          def clipScaledValue(outputScaledValue, outputRange):
              if (outputRange[0] < outputRange[1]):
                  return clipWhenLowerLimitIsLessThanHigher(outputScaledValue, outputRange)
              else:
                  return clipWhenLowerLimitIsGreaterThanHigherLimit(outputScaledValue, outputRange)
              end
          end

          def clipWhenLowerLimitIsGreaterThanHigherLimit(outputScaledValue, outputRange):
              if (outputScaledValue < outputRange[1]):
                  return outputRange[1]
              elif (outputScaledValue > outputRange[0]):
                  return outputRange[0]
              else:
                  return outputScaledValue
              end
          end

          def clipWhenLowerLimitIsLessThanHigher(outputScaledValue, outputRange):
              if (outputScaledValue < outputRange[0]):
                  return outputRange[0]
              elif (outputScaledValue > outputRange[1]):
                  return outputRange[1]
              else:
                  return outputScaledValue
              end
          end

          slope = computeSlope(rawRange, scaledRange)
          intercept = computeIntercept(slope, rawRange, scaledRange)
          scaledValue = slope * value + intercept
          return clipScaledValue(scaledValue, scaledRange)
      end

      def limit(value, range):
          return scale(value, range, range)
      end


  rq_init_comm_if_connected(9, "1")
  rq_init_comm_if_connected(2, "2")
  rq_init_comm_if_connected(3, "3")
  rq_init_comm_if_connected(4, "4")
  rq_print_connected_grippers()
  rq_gripper_communication_thread = run rq_gripper_communication()
  set_closed_norm(97.6470588235294, "1")
  set_open_norm(1.1764705882352942, "1")
  set_closed_mm(0.0, "1")
  set_open_mm(53.0, "1")
  set_closed_norm(100.0, "2")
  set_open_norm(0.0, "2")
  set_closed_mm(0.0, "2")
  set_open_mm(50.0, "2")
  set_closed_norm(100.0, "3")
  set_open_norm(0.0, "3")
  set_closed_mm(0.0, "3")
  set_open_mm(50.0, "3")
  set_closed_norm(100.0, "4")
  set_open_norm(0.0, "4")
  set_closed_mm(0.0, "4")
  set_open_mm(50.0, "4")
  rq_current_limit_enabled = False
  while(not rq_gripper_communication_thread_started):
      sleep(0.008)
  end
  # end: URCap Installation Node
  step_count_b1809ffc_a9dc_407a_9cc4_7bc2f4a6af46 = 0.0
  thread Step_Counter_Thread_37d5f412_1517_4c3d_9382_b16793093957():
    while (True):
      step_count_b1809ffc_a9dc_407a_9cc4_7bc2f4a6af46 = step_count_b1809ffc_a9dc_407a_9cc4_7bc2f4a6af46 + 1.0
      sync()
    end
  end
  run Step_Counter_Thread_37d5f412_1517_4c3d_9382_b16793093957()
  global AMR_Position=struct(position_identifier=0, x1=0, x2=0, y1=0, y2=0, theta1=0, theta2=0)
  global CAM_Pose=p[0,0,0,0,0,0]
  global CAM_Relation=""
  global CMD_Abort=  False
  global CMD_Clear=  False
  global CMD_Reset=  False
  global CMD_Start=  False
  global CMD_Suspend=  False
  global CMD_Unhold=  False
  global CMD_Unsuspend=  False
  global CNT_Rack_Output=0
  global FNC_Freedrive=  False
  global PRC_TubCounter=0
  global STP=0
  global easyPickCount_4=0
  global easyPickCount_6=0
  global easyPickCount_7=0
  global easyPickCount_8=0
  global easyPickCount_9=0
  global easyPickNoObj_4=0
  global easyPickNoObj_6=0
  global easyPickNoObj_7=0
  global easyPickNoObj_8=0
  global easyPickNoObj_9=0
  global easyPickParts_4=0
  global easyPickParts_6=0
  global easyPickParts_7=0
  global easyPickParts_8=0
  global easyPickParts_9=0
  global Dosing_time=0
  global TMR_Barcode=0
  global Container_mid_1_p=p[-.379239199143, -.127191311915, .299999999998, .000000000046, -.000000000021, -1.247199999994]
  global Container_mid_1_q=[-2.477408934449926, -1.2969853503591224, -1.875639182904262, -1.539621866126728, 1.5731943360401213, -2.8009955944022717]
  global trigger_otw_p=p[-.364831738276, -.163967193938, .343299997821, .000000000046, -.000000000020, -1.148401333327]
  global trigger_otw_q=[-2.378283213085033, -1.2994862387706814, -1.7634300687554951, -1.6493302004167063, 1.573123683454141, -2.8011223671816943]
  global Waypoint_54_p=p[.008800512419, -.547926542621, .402696567415, -.589884378425, -.007228654778, -.061268144704]
  global Waypoint_54_q=[-1.2044575850116175, -1.3416667741588135, -1.8272563219070435, -0.9884541195682068, 1.3621035814285278, -2.7712565104113978]
  global Waypoint_77_p=p[-.178371829612, -.433927395311, .368082383916, -.086593488055, .704679941724, -.007869906074]
  global Waypoint_77_q=[-1.265390698109762, -1.3355963987163086, -1.7944865226745605, -1.7402602634825648, 0.8780410885810852, -2.7713127771960657]
  global Waypoint_83_p=p[.008800512419, -.547926542621, .402696567415, -.589884378425, -.007228654778, -.061268144704]
  global Waypoint_83_q=[-1.2044575850116175, -1.3416667741588135, -1.8272563219070435, -0.9884541195682068, 1.3621035814285278, -2.7712565104113978]
  global Waypoint_84_p=p[-.178371829612, -.433927395311, .368082383916, -.086593488055, .704679941724, -.007869906074]
  global Waypoint_84_q=[-1.265390698109762, -1.3355963987163086, -1.7944865226745605, -1.7402602634825648, 0.8780410885810852, -2.7713127771960657]
  global Vial_above_1_p=p[.017105793010, -.652093028359, .184920586844, .000000000272, .000000000270, 1.564063451276]
  global Vial_above_1_q=[-1.3375440709712851, -1.9618096977868804, -1.4665759083780685, -1.2837941559171444, 1.5732503672317195, -4.47276330421513]
  global Vial_pick_poi_1_p=p[.017105792852, -.648922724010, .093307568731, .000000000271, .000000000270, 1.564063451276]
  global Vial_pick_poi_1_q=[-1.3366329456391917, -2.0375277831965413, -1.6071432798879028, -1.0675084332049813, 1.57309887265915, -4.471135348858068]
  global Waypoint_86_p=p[.019227646885, -.648669633640, .184920586950, .000000000000, .000000000000, .024063451426]
  global Waypoint_86_q=[-1.3331129109407733, -1.9540750545686123, -1.4775914902901128, -1.280581784992414, 1.5733500744865856, -2.928303704452631]
  global Waypoint_87_p=p[-.032361834699, -.348336136197, .391475576335, -.000008499254, .000014589902, -.004651426820]
  global Waypoint_87_q=[-1.2709335019096129, -1.1914598663441005, -1.708995335060501, -1.8117888533498316, 1.5729683532263925, -2.8379347397710237]
  global Vial_3FG_plac_1_p=p[-.031858676359, -.349402499566, .145301120695, .000000000000, .000000000000, .000000000000]
  global Vial_3FG_plac_1_q=[-1.2723975525801707, -1.252376585823825, -2.3128114007049496, -1.1470592278900167, 1.5730548099411423, -2.8414815174610535]
  global Waypoint_88_p=p[-.032361834699, -.348336136197, .391475576335, -.000008499254, .000014589902, -.004651426820]
  global Waypoint_88_q=[-1.2709335019096129, -1.1914598663441005, -1.708995335060501, -1.8117888533498316, 1.5729683532263925, -2.8379347397710237]
  global cap_dump_1_p=p[-.139168676487, -.420163541420, .146096395183, .000000000000, .000000000000, .000000000000]
  global cap_dump_1_q=[-1.584588644510994, -1.5093464179777323, -2.1118449369620347, -1.091059703602438, 1.5728943834877336, -3.154014906686923]
  global Waypoint_89_p=p[-.032361834699, -.348336136197, .391475576335, -.000008499254, .000014589902, -.004651426820]
  global Waypoint_89_q=[-1.2709335019096129, -1.1914598663441005, -1.708995335060501, -1.8117888533498316, 1.5729683532263925, -2.8379347397710237]
  global Vial_3FG_plac_2_p=p[-.031858676359, -.349402499566, .145301120695, .000000000000, .000000000000, .000000000000]
  global Vial_3FG_plac_2_q=[-1.2723975525801707, -1.252376585823825, -2.3128114007049496, -1.1470592278900167, 1.5730548099411423, -2.8414815174610535]
  global Waypoint_90_p=p[-.032361834699, -.348336136197, .391475576335, -.000008499254, .000014589902, -.004651426820]
  global Waypoint_90_q=[-1.2709335019096129, -1.1914598663441005, -1.708995335060501, -1.8117888533498316, 1.5729683532263925, -2.8379347397710237]
  global cap_dump_2_p=p[-.139168676487, -.420163541420, .146096395183, .000000000000, .000000000000, .000000000000]
  global cap_dump_2_q=[-1.584588644510994, -1.5093464179777323, -2.1118449369620347, -1.091059703602438, 1.5728943834877336, -3.154014906686923]
  global Waypoint_91_p=p[-.032361834699, -.348336136197, .391475576335, -.000008499254, .000014589902, -.004651426820]
  global Waypoint_91_q=[-1.2709335019096129, -1.1914598663441005, -1.708995335060501, -1.8117888533498316, 1.5729683532263925, -2.8379347397710237]
  global Vial_liq_abov_1_p=p[-.025303660977, -.338758622354, .426628485936, -1.315858642253, .800043520260, -.928295855026]
  global Vial_liq_abov_1_q=[-0.3789628187762659, -1.5149522957256814, -2.263045310974121, 0.7870649534412841, -0.750984017048971, -3.2237566153155726]
  global Vial_liq_pick_3_p=p[-.002660428945, -.335984893034, .159389832934, -1.150456778400, .673175527684, -1.010612657503]
  global Vial_liq_pick_3_q=[-0.3660772482501429, -1.4503649038127442, -2.4056053161621094, -1.994692941705221, 0.8039668202400208, -0.2508929411517542]
  global Vial_liq_pick_4_p=p[-.041402486291, -.356791603314, .125395323246, -1.143483969075, .651070210027, -.878721885453]
  global Vial_liq_pick_4_q=[-0.4426233705502476, -1.437252121513727, -2.551930962114307, -1.776528229806984, 0.6562026234073748, -0.43018811960029524]
  global Vial_liq_abov_2_p=p[-.025303660977, -.338758622354, .426628485936, -1.315858642253, .800043520260, -.928295855026]
  global Vial_liq_abov_2_q=[-0.3789628187762659, -1.5149522957256814, -2.263045310974121, 0.7870649534412841, -0.750984017048971, -3.2237566153155726]
  global Liquid_midway_1_p=p[.057575295009, -.583081747994, .306414980749, -1.351675548728, .120935756539, -.096908606303]
  global Liquid_midway_1_q=[-0.895174805318014, -1.7035466633238734, -2.380953073501587, 0.631549521083496, 0.7706599235534668, -2.9455552736865442]
  global shake_3_p=p[.057574880217, -.583085370269, .306422893466, -1.360996190983, -.155555042453, -.438136255921]
  global shake_3_q=[-0.8951800505267542, -1.7035466633238734, -2.380937099456787, 0.6315542894550782, 0.7706599235534669, -2.5394540616517496]
  global shake_4_p=p[.057581636113, -.583090570002, .306439684073, -1.308767904323, .368530312677, .214926493520]
  global shake_4_q=[-0.8951714674579065, -1.7035395107665003, -2.380906343460083, 0.6315504747578125, 0.7706480026245118, -3.3161255787892268]
  global drop_above_3_p=p[.268235025993, -.467784390499, .226219872376, -1.027832627524, -.430841408251, 1.004603115937]
  global drop_above_3_q=[-0.935645882283346, -1.6663371525206507, -2.4252893924713135, 0.41966931402172847, 1.8470635414123535, -3.4600217978106897]
  global drop_above_4_p=p[.219042229014, -.470775657081, .133754190740, -.313004595901, -.344395319364, 1.500564994056]
  global drop_above_4_q=[-1.0601594887284795, -1.70046459045642, -2.0799996233759863, -0.7243227230676759, 1.9429634314685202, -4.115129153870795]
  global liq_tran_3_p=p[.213067510942, -.469567035397, .100231043184, .251862243732, .217902579404, 1.592812335393]
  global liq_tran_3_q=[-0.7789645168037476, -1.822364827406652, -1.8643518410805573, -1.252158963840138, 1.3768134449520435, -3.9328333233290254]
  global drop_above_5_p=p[.219042229014, -.470775657081, .133754190740, -.313004595901, -.344395319364, 1.500564994056]
  global drop_above_5_q=[-1.0601594887284795, -1.70046459045642, -2.0799996233759863, -0.7243227230676759, 1.9429634314685202, -4.115129153870795]
  global Waypoint_92_p=p[.187119460405, -.493959476151, .133754190608, -.313004596540, -.344395317757, 1.500564993991]
  global Waypoint_92_q=[-1.1418328121400876, -1.7310553375189475, -2.033634768766424, -0.772026910513711, 1.958578934631971, -4.201588449364511]
  global liq_tran_4_p=p[.195957706507, -.493022614126, .100231042689, .160718757180, .109807038912, 1.525321508623]
  global liq_tran_4_q=[-0.881740380645474, -1.8244526267589851, -1.865100964490387, -1.1608866323693583, 1.4631433601076713, -3.973915130363038]
  global drop_above_6_p=p[.219042229014, -.470775657081, .133754190740, -.313004595901, -.344395319364, 1.500564994056]
  global drop_above_6_q=[-1.0601594887284795, -1.70046459045642, -2.0799996233759863, -0.7243227230676759, 1.9429634314685202, -4.115129153870795]
  global drop_above_7_p=p[.268235025993, -.467784390499, .226219872376, -1.027832627524, -.430841408251, 1.004603115937]
  global drop_above_7_q=[-0.935645882283346, -1.6663371525206507, -2.4252893924713135, 0.41966931402172847, 1.8470635414123535, -3.4600217978106897]
  global Liquid_midway_2_p=p[.057575295009, -.583081747994, .306414980749, -1.351675548728, .120935756539, -.096908606303]
  global Liquid_midway_2_q=[-0.895174805318014, -1.7035466633238734, -2.380953073501587, 0.631549521083496, 0.7706599235534668, -2.9455552736865442]
  global Vial_drop_abo_1_p=p[.000324902251, -.648569523142, .221894115667, -.873462921366, 1.165852672573, -1.482720593185]
  global Vial_drop_abo_1_q=[-1.0576906334721352, -2.393016994184633, -0.9236232851859159, -2.5729213042279273, 0.7903331288549689, -0.33286325848155585]
  global Vial_liq_drop_1_p=p[.001020867953, -.647659915585, .092915870838, -.834762611599, 1.081942994823, -1.540647900176]
  global Vial_liq_drop_1_q=[-1.0631954168193474, -2.4447642951220825, -1.128811017825127, -2.1983115491972294, 0.8130148661460634, -0.38984988696911316]
  global Vial_drop_abo_2_p=p[.000324902251, -.648569523142, .221894115667, -.873462921366, 1.165852672573, -1.482720593185]
  global Vial_drop_abo_2_q=[-1.0576906334721352, -2.393016994184633, -0.9236232851859159, -2.5729213042279273, 0.7903331288549689, -0.33286325848155585]
  global pick_cont_otw_p=p[-.479450777041, .284140798427, .125270103493, -.276792173670, 2.098433187454, -2.121256516887]
  global pick_cont_otw_q=[-2.891505066548503, -1.9549266300590151, -2.231827259067863, -1.6654960117542226, 0.020810842514162875, -0.4019392172601952]
  global Powder_wayp1_p=p[-.472820924474, .292439826233, .207418370237, -.137787250486, 2.177332259632, -2.152029714756]
  global Powder_wayp1_q=[-2.911134078210732, -1.90240864358569, -1.968768330510411, -2.500365101593811, 0.11427687110891149, 0.0958980389250167]
  global Waypoint_2_p=p[-.357612884176, -.251084817998, .212379799667, -.858181193174, 1.714832512191, -1.687547565568]
  global Waypoint_2_q=[-1.620834863369681, -1.8936194567376496, -1.9821394403832038, -2.4599791457905273, 0.6296693672615152, 0.07625365420707819]
  global Decapp_above_1_p=p[-.013480295948, -.359153355979, .266194408367, -.879653555922, 1.646336924805, -1.709111068605]
  global Decapp_above_1_q=[-0.9632157249872035, -2.0163405763031657, -1.5968194594157152, -2.6579215719847085, 1.251243398585566, 0.047906446502667066]
  global Decapp_place_2_p=p[-.013480295890, -.359153356055, .160907502384, -.879653554902, 1.646336919740, -1.709111066456]
  global Decapp_place_2_q=[-0.9633402410919709, -2.1541179572356635, -1.6937729380888573, -2.4232786481058053, 1.2517342187662468, 0.04818402956922263]
  global Decapp_above_2_p=p[-.013480295948, -.359153355979, .266194408367, -.879653555922, 1.646336924805, -1.709111068605]
  global Decapp_above_2_q=[-0.9632157249872035, -2.0163405763031657, -1.5968194594157152, -2.6579215719847085, 1.251243398585566, 0.047906446502667066]
  global Waypoint_78_p=p[-.051450028091, -.519555688329, .365718563414, -1.287302938145, 1.077637394477, -1.218524965834]
  global Waypoint_78_q=[-0.9214276262416012, -1.8899696965062578, -1.4939326452510562, -2.840015661555725, 0.5585157189668353, 0.033997638875617575]
  global Decap_above_p=p[-.031863883354, -.349974838955, .288042264213, .000000000000, .000000000000, .000000000000]
  global Decap_above_q=[-1.271900116540503, -1.1670201114602632, -1.989291655468758, -1.5559360538518163, 1.573255119759632, -2.842476569674073]
  global Decapp_p=p[-.031864263150, -.349974612700, .230259377740, .000000000000, .000000000000, .000000000000]
  global Decapp_q=[-1.2723555431601419, -1.1810456878410935, -2.1291754890757737, -1.4020263844320349, 1.5732701843074919, -2.842325632263757]
  global Cap_above_p=p[-.224192409203, -.629599568633, .257274081142, .000015605575, -.000015166009, -1.647823825902]
  global Cap_above_q=[-1.710642681834492, -1.9674285251810462, -1.2705185053146897, -1.4742193161331247, 1.573506065067499, -1.6347709465008595]
  global Cap_place_p=p[-.224189049846, -.629597879697, .041885651757, .000015605572, -.000015166011, -1.647823825903]
  global Cap_place_q=[-1.7111696563854295, -2.13979870939016, -1.5941008764912503, -0.978265561728648, 1.5732789016410962, -1.6336328794662904]
  global OP_PowderA2_p=p[.009371277507, -.409434369247, .294169017766, -.823281033205, 1.709410851243, -1.698303593897]
  global OP_PowderA2_q=[-0.9994544761745754, -2.1395254572673217, -1.3437567783153916, -2.8143375616690456, 1.2617899549595724, 0.019614613715634555]
  global OP_PowderA_ab_1_p=p[-.012145216791, -.363335041455, .315325728178, -.777135478411, 1.752984823781, -1.740925591659]
  global OP_PowderA_ab_1_q=[-1.01634425044037, -2.024785947780374, -1.4658894155189923, -2.8070189735738786, 1.3091674480404514, 0.020022086766872782]
  global OP_PowderA_pick_p=p[-.019989579300, -.367909055381, .180100616111, -.546164737600, 1.935964719000, -1.930057109666]
  global OP_PowderA_pick_q=[-1.1609156816971709, -2.238534265251247, -1.4969295335038062, -2.556223512058769, 1.4532886345781417, 0.020741051754957773]
  global OP_PowderA_ab_2_p=p[-.012145216791, -.363335041455, .315325728178, -.777135478411, 1.752984823781, -1.740925591659]
  global OP_PowderA_ab_2_q=[-1.01634425044037, -2.024785947780374, -1.4658894155189923, -2.8070189735738786, 1.3091674480404514, 0.020022086766872782]
  global Op_PowA_wP_p=p[-.173727579245, -.372934016396, .295116627479, -.972390492433, 1.540962074418, -1.548745344994]
  global Op_PowA_wP_q=[-1.1740587397768483, -1.865656321049359, -1.7426943793777419, -2.679427276872525, 0.8588908769087338, 0.017944699631825187]
  global Waypoint_1_p=p[-.451048883256, -.340589460864, .308223661552, .097058877504, .091048998701, -1.578386010942]
  global Waypoint_1_q=[-2.222400490437643, -1.7554131946959437, -1.398173213005066, -1.6564461193480433, 1.5042352676391602, -2.2106884161578577]
  global Spatula_otw_p=p[-.222059999126, -.318140885971, .425288233229, -.000441582509, -.000128175490, 3.034387645854]
  global Spatula_otw_q=[-1.827769217553847, -1.3054220991219179, -1.546249130536875, -1.8605379988907114, 1.573101813278913, -0.15105460523915326]
  global pick_spat_L_abv_p=p[.239059466375, -.067212518441, .280720723617, .000017217488, -.000484427718, 3.106837214660]
  global pick_spat_L_abv_q=[0.292765616142962, -0.8565557553273315, -2.140199892763044, -1.715349495646084, 1.573623142106424, 1.8984976776985687]
  global spat_L_pick_p=p[.242468789885, -.067301915011, .193171208067, .000017217488, -.000484427718, 3.106837214657]
  global spat_L_pick_q=[0.2867414378807389, -0.8600077002089179, -2.3629148016312627, -1.4891831672860159, 1.5737695566221115, 1.8933890858591198]
  global spat_L_lift_p=p[.245402002494, -.067432373551, .289049296496, .000017217490, -.000484427724, 3.106837214657]
  global spat_L_lift_q=[0.2834351187564135, -0.8798320076811592, -2.1119436738532986, -1.7203314352121302, 1.573588313403067, 1.8891054681654005]
  global spat_L_side_p=p[.247133573905, -.017633681797, .289062935631, .000017217490, -.000484427724, 3.106837214657]
  global spat_L_side_q=[0.49719173575848863, -0.8582398211168538, -2.1182130454788215, -1.735610316654931, 1.5735817737572706, 2.1028402698705397]
  global spat_L_up_p=p[.247135508752, -.017665230822, .397130746165, .000017217490, -.000484427724, 3.106837214657]
  global spat_L_up_q=[0.49854946074076967, -0.9346239623559676, -1.808280269374471, -1.969158816463132, 1.5731020084036995, 2.1031742024348157]
  global spat_M_up_p=p[.245495561680, -.112112573515, .420343789747, .000026293989, -.000477463067, 3.067686800858]
  global spat_M_up_q=[0.09017908059107435, -1.0134242235449396, -1.71728844067247, -1.9814399845077446, 1.573013686840385, 1.733759055129931]
  global spat_M_pick_p=p[.244673518506, -.111985070134, .192299022723, .000026293990, -.000477463072, 3.067686800901]
  global spat_M_pick_q=[0.08834054082534859, -0.9272467647495475, -2.3438023910348154, -1.4411029496965373, 1.5736983399628084, 1.7342144371718433]
  global spat_S_Up_1_p=p[.252087445596, -.159242094834, .423281604617, .000026293954, -.000477463070, 3.067686800855]
  global spat_S_Up_1_q=[-0.09804692328730358, -1.0862987822056382, -1.6788706463996483, -1.9470242450550348, 1.5730147401359813, 1.5455107082823842]
  global spat_S_Pick_1_p=p[.245377020686, -.158668022535, .192285730279, .000026293985, -.000477463062, 3.067686800840]
  global spat_S_Pick_1_q=[-0.10087203759495189, -1.011188488703386, -2.311978084495874, -1.3890267520590838, 1.5735990551056096, 1.5450562970948172]
  global spat_S_Up_2_p=p[.252087445596, -.159242094834, .423281604617, .000026293954, -.000477463070, 3.067686800855]
  global spat_S_Up_2_q=[-0.09804692328730358, -1.0862987822056382, -1.6788706463996483, -1.9470242450550348, 1.5730147401359813, 1.5455107082823842]
  global spat_flatM_up_p=p[.229022666361, -.211442909333, .418634047126, .000026293953, -.000477463083, 3.067686800888]
  global spat_flatM_up_q=[-0.30183372580416545, -1.1157042924275036, -1.6775646144685776, -1.9189678841796578, 1.5730340557943228, 1.341766142011193]
  global spat_flatM_pick_p=p[.241028983327, -.208057297586, .192270533170, .000026293950, -.000477463079, 3.067686800885]
  global spat_flatM_pick_q=[-0.2805687960562633, -1.1003763929487214, -2.271431297337675, -1.3404236887924883, 1.5734924238720627, 1.3653813047742556]
  global spat_flatS_up_p=p[.237651953780, -.253943828614, .403961222825, .000026293950, -.000477463092, 3.067686800841]
  global spat_flatS_up_q=[-0.42363550926974103, -1.1939944599502539, -1.6745915127240307, -1.843675057902054, 1.5731001874678698, 1.220082820532415]
  global spat_flatS_pick_p=p[.241325662334, -.251726327528, .192256842740, .000026293947, -.000477463087, 3.067686800841]
  global spat_flatS_pick_q=[-0.4144907797170738, -1.1967447109013012, -2.21926362252748, -1.2962499335425761, 1.5733885098427622, 1.2314402238866728]
  global spat_S_pick_p=p[.238158866340, -.157926795425, .192632100345, .000026293989, -.000477463069, 3.067686800857]
  global spat_S_pick_q=[-0.10084756991493293, -0.9881392730064915, -2.3204232610157494, -1.403630829593915, 1.5736254260650586, 1.5450653591083503]
  global spat_S_up_p=p[.244260523725, -.164466690315, .417087579736, .000026293988, -.000477463072, 3.067686800857]
  global spat_S_up_q=[-0.12101499604198729, -1.0718307017854336, -1.7023391702814736, -1.938028805938881, 1.573044424728474, 1.5226045951991447]
  global spat_S_Up_3_p=p[.252087445596, -.159242094834, .423281604617, .000026293954, -.000477463070, 3.067686800855]
  global spat_S_Up_3_q=[-0.09804692328730358, -1.0862987822056382, -1.6788706463996483, -1.9470242450550348, 1.5730147401359813, 1.5455107082823842]
  global spat_S_Pick_2_p=p[.245377020686, -.158668022535, .192285730279, .000026293985, -.000477463062, 3.067686800840]
  global spat_S_Pick_2_q=[-0.10087203759495189, -1.011188488703386, -2.311978084495874, -1.3890267520590838, 1.5735990551056096, 1.5450562970948172]
  global spat_S_Up_4_p=p[.252087445596, -.159242094834, .423281604617, .000026293954, -.000477463070, 3.067686800855]
  global spat_S_Up_4_q=[-0.09804692328730358, -1.0862987822056382, -1.6788706463996483, -1.9470242450550348, 1.5730147401359813, 1.5455107082823842]
  global PosA_up_p=p[.016801192651, -.634607931192, .234972649145, -1.090660933959, 1.404791542935, -1.413645191218]
  global PosA_up_q=[-1.0269853941957567, -2.5566815932087046, -0.7524196965257657, -2.981505396440104, 0.8113680441070815, 0.02148045637209592]
  global PosA_pick_p=p[.015038978729, -.636805282702, .098001171702, -1.090660933960, 1.404791542941, -1.413645191214]
  global PosA_pick_q=[-1.030538681681108, -2.6868026737636344, -0.8591268496433386, -2.7445819191995, 0.8086593798745287, 0.021358164952170952]
  global trigger_otw_2_p=p[-.364831738276, -.163967193938, .343299997821, .000000000046, -.000000000020, -1.148401333327]
  global trigger_otw_2_q=[-2.378283213085033, -1.2994862387706814, -1.7634300687554951, -1.6493302004167063, 1.573123683454141, -2.8011223671816943]
  global Postions_otw_p=p[-.010896578244, -.533368729951, .288851175116, -1.233738470894, 1.195331112012, -1.207314088469]
  global Postions_otw_q=[-0.898791023514228, -2.078490033037677, -1.4499891355755317, -2.7624416226992476, 0.6570218891920963, 0.02136606178275929]
  global spat_S_Up_5_p=p[.252087445596, -.159242094834, .423281604617, .000026293954, -.000477463070, 3.067686800855]
  global spat_S_Up_5_q=[-0.09804692328730358, -1.0862987822056382, -1.6788706463996483, -1.9470242450550348, 1.5730147401359813, 1.5455107082823842]
  global spat_S_Pick_3_p=p[.245377020686, -.158668022535, .192285730279, .000026293985, -.000477463062, 3.067686800840]
  global spat_S_Pick_3_q=[-0.10087203759495189, -1.011188488703386, -2.311978084495874, -1.3890267520590838, 1.5735990551056096, 1.5450562970948172]
  global spat_S_Up_6_p=p[.252087445596, -.159242094834, .423281604617, .000026293954, -.000477463070, 3.067686800855]
  global spat_S_Up_6_q=[-0.09804692328730358, -1.0862987822056382, -1.6788706463996483, -1.9470242450550348, 1.5730147401359813, 1.5455107082823842]
  global spat_S_Up_7_p=p[.252087445596, -.159242094834, .423281604617, .000026293954, -.000477463070, 3.067686800855]
  global spat_S_Up_7_q=[-0.09804692328730358, -1.0862987822056382, -1.6788706463996483, -1.9470242450550348, 1.5730147401359813, 1.5455107082823842]
  global spat_S_Pick_4_p=p[.245377020686, -.158668022535, .192285730279, .000026293985, -.000477463062, 3.067686800840]
  global spat_S_Pick_4_q=[-0.10087203759495189, -1.011188488703386, -2.311978084495874, -1.3890267520590838, 1.5735990551056096, 1.5450562970948172]
  global spat_S_Up_8_p=p[.252087445596, -.159242094834, .423281604617, .000026293954, -.000477463070, 3.067686800855]
  global spat_S_Up_8_q=[-0.09804692328730358, -1.0862987822056382, -1.6788706463996483, -1.9470242450550348, 1.5730147401359813, 1.5455107082823842]
  global PosB_up_p=p[.239472634782, -.492481416782, .220767759213, -1.233738470883, 1.195331111998, -1.207314088469]
  global PosB_up_q=[-0.5800230603397054, -2.4076296700885997, -1.0699783327330836, -2.8116344407747427, 0.9750472858169287, 0.017627507888886562]
  global PosB_pick_p=p[.240630296955, -.494558620171, .096392895280, -1.233740573549, 1.195309876041, -1.207293779132]
  global PosB_pick_q=[-0.5816146260408139, -2.553273721769836, -1.1376320925804277, -2.5983292591462153, 0.9740936784345416, 0.017625262979849232]
  global PosC_up_p=p[.241566602786, -.359249123455, .230260583862, -1.233738470888, 1.195331111997, -1.207314088449]
  global PosC_up_q=[-0.39573787962534546, -2.2019009616581497, -1.4115270142506517, -2.675987785326166, 1.160180741930842, 0.01687917643039505]
  global PosC_pick_p=p[.240633854030, -.361553124916, .093979792658, -1.233738470878, 1.195331111997, -1.207314088469]
  global PosC_pick_q=[-0.39992427526118757, -2.386042391328985, -1.4894374567278712, -2.414022930893381, 1.1566786195951169, 0.01712017454263659]
  global Pow_decap_up_p=p[-.017556487132, -.367519866742, .275835445416, -.605635182849, 1.892518157522, -1.890848751165]
  global Pow_decap_up_q=[-1.1272088681128203, -2.1173924123331025, -1.4250048354055203, -2.7485980486387676, 1.4193896902217862, 0.023247957637719453]
  global pow_decap_place_p=p[-.020433194420, -.368310202914, .161281291611, -.605635182838, 1.892518157522, -1.890848751163]
  global pow_decap_place_q=[-1.132360890531647, -2.2521863255983092, -1.5302136899970318, -2.5086176644751683, 1.4149282844269635, 0.02347140074572661]
  global Decap_up_p=p[-.018339217391, -.367674469480, .249553854268, -.546164737599, 1.935964719000, -1.930057109666]
  global Decap_up_q=[-1.158124747223252, -2.1569920012936787, -1.4340832185069745, -2.7006032680036753, 1.4556626828962336, 0.02060977878679182]
  global Decap_pick_p=p[-.020429098827, -.367971872627, .161604333799, -.546164737600, 1.935964719000, -1.930057109666]
  global Decap_pick_q=[-1.161653098289774, -2.263509236689538, -1.5087211318402236, -2.519459740767391, 1.452646640403743, 0.02077912034002202]
  global spat_S_Up_9_p=p[.252087445596, -.159242094834, .423281604617, .000026293954, -.000477463070, 3.067686800855]
  global spat_S_Up_9_q=[-0.09804692328730358, -1.0862987822056382, -1.6788706463996483, -1.9470242450550348, 1.5730147401359813, 1.5455107082823842]
  global spat_S_Pick_5_p=p[.245377020686, -.158668022535, .192285730279, .000026293985, -.000477463062, 3.067686800840]
  global spat_S_Pick_5_q=[-0.10087203759495189, -1.011188488703386, -2.311978084495874, -1.3890267520590838, 1.5735990551056096, 1.5450562970948172]
  global spat_S_Up_10_p=p[.252087445596, -.159242094834, .423281604617, .000026293954, -.000477463070, 3.067686800855]
  global spat_S_Up_10_q=[-0.09804692328730358, -1.0862987822056382, -1.6788706463996483, -1.9470242450550348, 1.5730147401359813, 1.5455107082823842]
  global Cap_Pos1_up_p=p[-.009204590651, -.630414532143, .209553215594, .000015605636, -.000015165972, -1.647823825918]
  global Cap_Pos1_up_q=[-1.3712235360848153, -1.8956436160717116, -1.4937179908129403, -1.3227667547680468, 1.5734078303557693, -1.294583528806303]
  global Cap_pos1_p=p[-.009202676635, -.630420568421, .169124041327, .000015605637, -.000015165972, -1.647823825918]
  global Cap_pos1_q=[-1.3713472255781163, -1.9233675297983162, -1.5632855513360973, -1.2254750650219144, 1.573366428933177, -1.2943660310427454]
  global Cap_Pos2_up_p=p[.211716053312, -.494057775376, .215280069366, .000015605634, -.000015165975, -1.647823825915]
  global Cap_Pos2_up_q=[-0.9145242936692304, -1.674696899505042, -1.7522162453415309, -1.2851708271213624, 1.5732187144557628, -0.8372657504386876]
  global Cap_Pos2_p=p[.212489912868, -.496566704351, .174147693321, .000015605636, -.000015165975, -1.647823825915]
  global Cap_Pos2_q=[-0.9164207524863208, -1.713567851985026, -1.8189683536262713, -1.1795477490971313, 1.5731464491112233, -0.8388186043721344]
  global Cap_Pos3_up_p=p[.215414026072, -.362498267015, .204704869421, .000015605620, -.000015165977, -1.647823825911]
  global Cap_Pos3_up_q=[-0.7126949721702758, -1.3944102858194336, -2.0491785338653417, -1.268480216466319, 1.5731602525658304, -0.6347529509142049]
  global Cap_pos3_p=p[.215414769079, -.362497999431, .173969495144, .000015605637, -.000015165975, -1.647823825916]
  global Cap_pos3_q=[-0.7128543668961971, -1.4224209260451453, -2.1096401714367516, -1.1800078429832341, 1.573077069822543, -0.6346164729408441]
  global Dosing_time_is_counting=False
  global TMR_Barcode_is_counting=False
  thread Timer_Thread():
    while (True):
      if (Dosing_time_is_counting):
        Dosing_time = Dosing_time + get_steptime()
      end
      if (TMR_Barcode_is_counting):
        TMR_Barcode = TMR_Barcode + get_steptime()
      end
      sync()
    end
  end
  run Timer_Thread()
  def Sub_Vision_V18():
    $ 817 "Sub_Vision_V18" "noBreak"
    $ 818 "PreSettings"
    $ 819 "CAM_LM_Detected≔ False "
    global CAM_LM_Detected=  False
    $ 820 "CAM_Captures≔0"
    global CAM_Captures=0
    $ 821 "CAM_Pose≔p[0,0,0,0,0,0]"
    global CAM_Pose=p[0,0,0,0,0,0]
    $ 822 "CAM_LM_Refinmnt≔ False "
    global CAM_LM_Refinmnt=  False
    $ 823 "CAM_LM_Refined≔ False "
    global CAM_LM_Refined=  False
    $ 824 "CAM_LM_Deviatn≔p[0,0,0,0,0,0]"
    global CAM_LM_Deviatn=p[0,0,0,0,0,0]
    $ 825 "CAM_LM_ID≔0"
    global CAM_LM_ID=0
    $ 826 "CAM_Done≔ False "
    global CAM_Done=  False
    $ 827 "CAM_CNT_Obj≔0"
    global CAM_CNT_Obj=0
    $ 828 "CAM_Result = []"
    CAM_Result = []
    $ 829 "OBJ_Detected≔ False "
    global OBJ_Detected=  False
    $ 830 "FRM_Reference≔p[0,0,0,0,0,0]"
    global FRM_Reference=p[0,0,0,0,0,0]
    $ 831 "'=========='"
    # '=========='
    $ 832 "Switch Action"
    switch_1 = Action
    $ 833 "Case 13"
    if (13 == switch_1):
    elif (15 == switch_1):
      $ 951 "Case 15"
    elif (131 == switch_1):
      $ 997 "Case 131"
      $ 998 "Read (SensoPart)"
      $ 999 "Action_Info≔'search for landmark'"
      global Action_Info="search for landmark"
      $ 1000 "CAM_LM≔CAM_LMs[4]"
      global CAM_LM=CAM_LMs[4]
      $ 1001 "CAM_Relation≔CAM_LM.capture_relation"
      global CAM_Relation=CAM_LM.capture_relation
      $ 1002 "go to capture pose"
      $ 1005 "If ITM_ID≟1 and JIG≟7"
      if (ITM_ID == 1  and  JIG == 7):
        $ 1006 "PSE_T≔uLM_Cap_SSRack"
        global PSE_T=uLM_Cap_SSRack
      else:
        $ 1007 "ElseIf ITM_ID≟5 and JIG≟7"
        if (ITM_ID == 5  and  JIG == 7):
          $ 1008 "PSE_T≔FRM_Cap_SSRack"
          global PSE_T=FRM_Cap_SSRack
        else:
          $ 1011 "ElseIf ITM_ID≟1 and JIG≟15"
          if (ITM_ID == 1 and JIG == 15):
            $ 1012 "MoveJ"
            $ 1013 "Container_mid_1" "breakAfter"
            movej(get_inverse_kin(Container_mid_1_p, qnear=Container_mid_1_q), a=1.3962634015954636, v=1.0471975511965976, r=0.05)
            $ 1015 "PSE_T≔FRM_Container_const"
            global PSE_T=p[-0.5003348223692186,0.35061804815168285,0.41579001388808423,-5.092943187272062E-5,1.0145185065363121E-4,-2.764319258713288]
          else:
            $ 1016 "ElseIf ITM_ID≟1 and JIG≟21"
            if (ITM_ID == 1 and JIG == 21):
              $ 1017 "PSE_T≔FRM_PoTS_const"
              global PSE_T=p[-0.5306792777448894,-0.11733736113273928,0.4723291514857741,-1.2750528643267135E-5,1.622694849249343E-6,-2.208498084105121]
            else:
              $ 1018 "ElseIf ITM_ID≟1 and JIG≟17"
              if (ITM_ID == 1 and JIG == 17):
                $ 1019 "MoveJ"
                $ 1020 "trigger_otw" "breakAfter"
                movej(get_inverse_kin(trigger_otw_p, qnear=trigger_otw_q), a=1.3962634015954636, v=1.0471975511965976, r=0.05)
                $ 1021 "PSE_T≔FRM_weigh_scale_const"
                global PSE_T=p[-0.3552030492367321,0.06852934966463993,0.4723405535118315,-1.0342323845904682E-4,-1.3726098069249118E-5,-2.169178331189411]
              end
            end
          end
        end
      end
      $ 1022 "do_transition(PSE_T, keep_rxry=False)"
      do_transition(PSE_T, keep_rxry=False)
      $ 1023 "Set"
      set_tcp(p[0.0,0.0,0.161,3.1415,0.0,0.0])
      $ 1024 "MoveJ"
      $ 1025 "PSE_T" "breakAfter"
      movej(PSE_T, a=1.3962634015954636, v=1.7453292519943295)
      $ 1026 "CAM_Pose≔get_actual_tcp_pose()"
      global CAM_Pose= get_actual_tcp_pose ()
      $ 1027 "Loop  not CAM_Done and  not ERROR.FLAG and  not CMD_Stop"
      while (  not  CAM_Done  and    not  ERROR.FLAG  and    not  CMD_Stop):
        $ 1028 "adjust capture pose"
        $ 1029 "If CAM_LM_Detected and CAM_LM_Refinmnt"
        if (CAM_LM_Detected  and  CAM_LM_Refinmnt):
          $ 1030 "PSE_T≔p[0,0,0.300,0,0,0]"
          global PSE_T=p[0,0,0.300,0,0,0]
          $ 1031 "CAM_Pose≔PSE_T"
          global CAM_Pose=PSE_T
          $ 1032 "If  not is_reachable(FRM_Reference,[PSE_T])"
          if (  not  is_reachable(FRM_Reference,[PSE_T])):
            $ 1033 "Error"
            $ 1034 "set_error(ERROR_POSE_NOT_REACHABLE)"
            set_error(ERROR_POSE_NOT_REACHABLE)
          end
          $ 1035 "If  not ERROR.FLAG"
          if (  not  ERROR.FLAG):
            $ 1036 "MoveJ"
            $ 1037 "PSE_T" "breakAfter"
            set_tcp(p[0.0,0.0,0.161,0.0,0.0,0.0])
            movej(pose_trans(FRM_Reference, PSE_T), a=0.8726646259971648, v=1.3962634015954636)
            $ 1038 "CAM_LM_Refined≔ True "
            global CAM_LM_Refined=  True
          end
        else:
          $ 1039 "ElseIf  not CAM_LM_Detected and CAM_Captures>0"
          if (  not  CAM_LM_Detected  and  CAM_Captures>0):
            $ 1040 "MoveL"
            $ 1041 "If FRM_Reference≟p[0,0,0,0,0,0]"
            if (FRM_Reference == p[0,0,0,0,0,0]):
              $ 1042 "PSE_T≔get_random_pose(pose_ref=CAM_Pose, mode='cubic', range_max=[0.150,0.150,0.015])"
              global PSE_T=get_random_pose(pose_ref=CAM_Pose, mode="cubic", range_max=[0.150,0.150,0.015])
            else:
              $ 1047 "Else" "noBreak"
              $ 1048 "PSE_T≔get_random_pose(pose_ref=CAM_Pose, mode='rotation', range_max=[10,10,0])"
              global PSE_T=get_random_pose(pose_ref=CAM_Pose, mode="rotation", range_max=[10,10,0])
              $ 1049 "CAM_LM_Refined≔ True "
              global CAM_LM_Refined=  True
            end
            $ 1050 "If get_inverse_kin_has_solution(pose_trans(FRM_Reference, PSE_T))"
            if (get_inverse_kin_has_solution( pose_trans (FRM_Reference, PSE_T))):
              $ 1051 "Comment"
              # Comment
              $ 1052 "PSE_T" "breakAfter"
              set_tcp(p[0.0,0.0,0.161,3.1415,0.0,0.0])
              movel(pose_trans(FRM_Reference, PSE_T), a=0.03, v=0.05)
            else:
              $ 1053 "Else" "noBreak"
              $ 1054 "'If random pose is out of reach, set the initial cam pose'"
              # 'If random pose is out of reach, set the initial cam pose'
              $ 1055 "PSE_T≔CAM_Pose"
              global PSE_T=CAM_Pose
            end
          end
        end
        $ 1056 "Wait: 2.0"
        sleep(2.0)
        $ 1057 "trigger"
        $ 1058 "If ITM_ID≟1 and JIG≟7"
        if (ITM_ID == 1  and  JIG == 7):
          # begin: URCap Program Node
          #   Source: SensoPart VISOR Robotic, 2.0.6, SensoPart Industriesensorik GmbH
          #   Type: VISOR Trigger
          $ 1059 "# 1 VISOR Trigger"
          visor_changeJob(1, "Landmark_INVITE_2", 6000)
          visor_trigger(1, 6000, "arm")
          # end: URCap Program Node
        else:
          $ 1060 "ElseIf ITM_ID≟5 and JIG≟7"
          if (ITM_ID == 5  and  JIG == 7):
            # begin: URCap Program Node
            #   Source: SensoPart VISOR Robotic, 2.0.6, SensoPart Industriesensorik GmbH
            #   Type: VISOR Trigger
            $ 1061 "# 1 VISOR Trigger"
            visor_changeJob(1, "Landmark_INVITE_2", 6000)
            visor_trigger(1, 6000, "arm")
            # end: URCap Program Node
          else:
            $ 1062 "ElseIf ITM_ID≟13 and JIG≟7"
            if (ITM_ID == 13  and  JIG == 7):
              # begin: URCap Program Node
              #   Source: SensoPart VISOR Robotic, 2.0.6, SensoPart Industriesensorik GmbH
              #   Type: VISOR Trigger
              $ 1063 "# 1 VISOR Trigger"
              visor_changeJob(1, "Landmark_INVITE_2", 6000)
              visor_trigger(1, 6000, "arm")
              # end: URCap Program Node
            else:
              $ 1064 "ElseIf ITM_ID≟1 and JIG≟15"
              if (ITM_ID == 1 and JIG == 15):
                # begin: URCap Program Node
                #   Source: SensoPart VISOR Robotic, 2.0.6, SensoPart Industriesensorik GmbH
                #   Type: VISOR Trigger
                $ 1065 "# 1 VISOR Trigger"
                visor_changeJob(1, "QR_box", 6000)
                visor_trigger(1, 6000, "arm")
                # end: URCap Program Node
              else:
                $ 1066 "ElseIf ITM_ID≟1 and JIG≟21"
                if (ITM_ID == 1 and JIG == 21):
                  # begin: URCap Program Node
                  #   Source: SensoPart VISOR Robotic, 2.0.6, SensoPart Industriesensorik GmbH
                  #   Type: VISOR Trigger
                  $ 1067 "# 1 VISOR Trigger"
                  visor_changeJob(1, "PoTS", 6000)
                  visor_trigger(1, 6000, "arm")
                  # end: URCap Program Node
                else:
                  $ 1068 "ElseIf ITM_ID≟1 and JIG≟17"
                  if (ITM_ID == 1 and JIG == 17):
                    # begin: URCap Program Node
                    #   Source: SensoPart VISOR Robotic, 2.0.6, SensoPart Industriesensorik GmbH
                    #   Type: VISOR Trigger
                    $ 1069 "# 1 VISOR Trigger"
                    visor_changeJob(1, "Weigh_target", 6000)
                    visor_trigger(1, 6000, "arm")
                    # end: URCap Program Node
                  end
                end
              end
            end
          end
        end
        $ 1073 "TM_3D_Found≔visor_partsFound(1)"
        global TM_3D_Found= visor_partsFound (1)
        $ 1074 "If TM_3D_Found>0"
        if (TM_3D_Found>0):
          $ 1075 "CAM_LM_Detected≔ True "
          global CAM_LM_Detected=  True
          $ 1076 "CAM_Captures≔0"
          global CAM_Captures=0
        else:
          $ 1077 "Else" "noBreak"
          $ 1078 "CAM_LM_Detected≔ False "
          global CAM_LM_Detected=  False
          $ 1079 "CAM_Captures≔CAM_Captures+1"
          global CAM_Captures=CAM_Captures+1
        end
        $ 1084 "result"
        $ 1085 "If CAM_LM_Detected"
        if (CAM_LM_Detected):
          $ 1086 "If (CAM_LM_Refinmnt and CAM_LM_Refined) or  not CAM_LM_Refinmnt"
          if ((CAM_LM_Refinmnt  and  CAM_LM_Refined)  or    not  CAM_LM_Refinmnt):
            $ 1144 "If ITM_ID≟1 and JIG≟7"
            if (ITM_ID == 1  and  JIG == 7):
              $ 1145 "CAM_LM_SSRack≔visor_getPose3d(1, 0)"
              global CAM_LM_SSRack= visor_getPose3d (1, 0)
            else:
              $ 1146 "ElseIf ITM_ID≟5 and JIG≟7"
              if (ITM_ID == 5  and  JIG == 7):
                $ 1147 "CAM_LM_SSRack≔visor_getPose3d(1, 0)"
                global CAM_LM_SSRack= visor_getPose3d (1, 0)
              else:
                $ 1150 "ElseIf ITM_ID≟1 and JIG≟15"
                if (ITM_ID == 1 and JIG == 15):
                  $ 1151 "CAM_LM_cont≔visor_getPose3d(1, 0)"
                  global CAM_LM_cont= visor_getPose3d (1, 0)
                  $ 1152 "Trigger≔get_actual_tcp_pose()"
                  global Trigger= get_actual_tcp_pose ()
                else:
                  $ 1153 "ElseIf ITM_ID≟1 and JIG≟21"
                  if (ITM_ID == 1 and JIG == 21):
                    $ 1154 "CAM_LM_cont≔visor_getPose3d(1, 0)"
                    global CAM_LM_cont= visor_getPose3d (1, 0)
                    $ 1155 "Trigger≔get_actual_tcp_pose()"
                    global Trigger= get_actual_tcp_pose ()
                  else:
                    $ 1156 "ElseIf ITM_ID≟1 and JIG≟17"
                    if (ITM_ID == 1 and JIG == 17):
                      $ 1157 "CAM_LM_cont≔visor_getPose3d(1, 0)"
                      global CAM_LM_cont= visor_getPose3d (1, 0)
                      $ 1158 "Trigger≔get_actual_tcp_pose()"
                      global Trigger= get_actual_tcp_pose ()
                    end
                  end
                end
              end
            end
            $ 1159 "CAM_Done≔ True "
            global CAM_Done=  True
          end
        else:
          $ 1160 "ElseIf  not CAM_LM_Detected and CAM_Captures<CAM_PRM_Retries"
          if (  not  CAM_LM_Detected  and  CAM_Captures<CAM_PRM_Retries):
            $ 1161 "CAM_LM_Refined≔ False "
            global CAM_LM_Refined=  False
          else:
            $ 1162 "ElseIf CAM_Captures≥CAM_PRM_Retries"
            if (CAM_Captures >= CAM_PRM_Retries):
              $ 1163 "CAM_Done≔ True "
              global CAM_Done=  True
              $ 1164 "Error"
              $ 1165 "set_error(ERROR_NO_LANDMARK)"
              set_error(ERROR_NO_LANDMARK)
            end
          end
        end
      end
    elif (151 == switch_1):
      $ 1166 "Case 151"
      $ 1167 "Detect (SensoPart)"
      $ 1168 "go to capture pose"
      $ 1169 "FRM_Reference≔FRM_Cap_SSRack"
      global FRM_Reference=FRM_Cap_SSRack
      $ 1170 "PSE_T≔p[0,0,-0.00,0,0,0]"
      global PSE_T=p[0,0,-0.00,0,0,0]
      $ 1171 "do_transition(pose_trans(FRM_Reference, PSE_T), keep_rxry=False)"
      do_transition( pose_trans (FRM_Reference, PSE_T), keep_rxry=False)
      $ 1172 "JNT_Q≔get_actual_joint_positions()"
      global JNT_Q= get_actual_joint_positions ()
      $ 1173 "JNT_Q≔[JNT_Q[0], JNT_Q[1], JNT_Q[2], JNT_Q[3], JNT_Q[4], 0]"
      global JNT_Q=[JNT_Q[0], JNT_Q[1], JNT_Q[2], JNT_Q[3], JNT_Q[4], 0]
      $ 1174 "Set"
      set_tcp(p[0.0,0.0,0.161,3.1415,0.0,0.0])
      $ 1175 "movej(get_inverse_kin(pose_trans(FRM_Reference, PSE_T), qnear=JNT_Q))"
      movej(get_inverse_kin( pose_trans (FRM_Reference, PSE_T), qnear=JNT_Q))
      $ 1176 "CAM_Pose≔pose_trans(pose_inv(FRM_Reference), get_actual_tcp_pose())"
      global CAM_Pose= pose_trans ( pose_inv (FRM_Reference),  get_actual_tcp_pose ())
      $ 1177 "Loop  not CAM_Done and  not ERROR.FLAG and  not CMD_Stop"
      while (  not  CAM_Done  and    not  ERROR.FLAG  and    not  CMD_Stop):
        $ 1178 "If  not OBJ_Detected and CAM_Captures>0"
        if (  not  OBJ_Detected  and  CAM_Captures>0):
          $ 1179 "MoveL"
          $ 1180 "If FRM_Reference≟p[0,0,0,0,0,0]"
          if (FRM_Reference == p[0,0,0,0,0,0]):
            $ 1182 "PSE_T≔get_random_pose(pose_ref=CAM_Pose, mode='rotation', range_max=[15,15,0])"
            global PSE_T=get_random_pose(pose_ref=CAM_Pose, mode="rotation", range_max=[15,15,0])
          else:
            $ 1183 "Else" "noBreak"
            $ 1184 "PSE_T≔get_random_pose(pose_ref=CAM_Pose, mode='rotation', range_max=[10,10,0])"
            global PSE_T=get_random_pose(pose_ref=CAM_Pose, mode="rotation", range_max=[10,10,0])
          end
          $ 1185 "If get_inverse_kin_has_solution(pose_trans(FRM_Reference, PSE_T))"
          if (get_inverse_kin_has_solution( pose_trans (FRM_Reference, PSE_T))):
            $ 1186 "PSE_T" "breakAfter"
            set_tcp(p[0.0,0.0,0.161,3.1415,0.0,0.0])
            movel(pose_trans(FRM_Reference, PSE_T), a=0.03, v=0.05)
          else:
            $ 1187 "Else" "noBreak"
            $ 1188 "'If random pose is out of reach, set the initial cam pose'"
            # 'If random pose is out of reach, set the initial cam pose'
            $ 1189 "PSE_T≔CAM_Pose"
            global PSE_T=CAM_Pose
            $ 1190 "PSE_T" "breakAfter"
            set_tcp(p[0.0,0.0,0.161,3.1415,0.0,0.0])
            movel(pose_trans(FRM_Reference, PSE_T), a=0.03, v=0.05)
          end
        end
        $ 1191 "Wait: 0.5"
        sleep(0.5)
        $ 1192 "Set"
        set_tcp(p[0.0,0.0,0.161,3.1415,0.0,0.0])
        # begin: URCap Program Node
        #   Source: SensoPart VISOR Robotic, 2.0.6, SensoPart Industriesensorik GmbH
        #   Type: VISOR Trigger
        $ 1193 "# 1 VISOR Trigger"
        visor_changeJob(1, "Object Detection Single", 6000)
        visor_trigger(1, 6000, "arm")
        # end: URCap Program Node
        $ 1194 "If visor_isResponseOk(1)"
        if ( visor_isResponseOk (1)):
          $ 1195 "CAM_CNT_Obj≔visor_partsFound(1)"
          global CAM_CNT_Obj= visor_partsFound (1)
          $ 1196 "CAM_OBJ_Pose≔visor_getPose3d(1, 0)"
          global CAM_OBJ_Pose= visor_getPose3d (1, 0)
          $ 1197 "If CAM_CNT_Obj>0"
          if (CAM_CNT_Obj>0):
            $ 1198 "CAM_OBJ_Color≔visor_getAdditionalData(1, 0)"
            global CAM_OBJ_Color= visor_getAdditionalData (1, 0)
            $ 1199 "CAM_DetectScore≔to_num(visor_getAdditionalData(1, 1))/1000"
            global CAM_DetectScore=to_num( visor_getAdditionalData (1, 1))/1000
            $ 1200 "OBJ_Detected≔ True "
            global OBJ_Detected=  True
          end
        else:
          $ 1201 "Else" "noBreak"
          $ 1202 "CAM_Captures≔CAM_Captures+1"
          global CAM_Captures=CAM_Captures+1
        end
        $ 1203 "If OBJ_Detected"
        if (OBJ_Detected):
          $ 1204 "Get object data"
          $ 1205 "PRC_CntDetect≔0"
          global PRC_CntDetect=0
          $ 1206 "Loop PRC_CntDetect<CAM_CNT_Obj"
          while (PRC_CntDetect<CAM_CNT_Obj):
            $ 1207 "get object and jig number"
            $ 1208 "If ITM_ID≟1 and JIG≟7"
            if (ITM_ID == 1  and  JIG == 7):
              $ 1209 "FRM_Reference≔FRM_Cap_SSRack"
              global FRM_Reference=FRM_Cap_SSRack
            else:
              $ 1210 "ElseIf ITM_ID≟5 and JIG≟7"
              if (ITM_ID == 5  and  JIG == 7):
                $ 1211 "FRM_Reference≔uLM_Cap_SSRack"
                global FRM_Reference=uLM_Cap_SSRack
              end
            end
            $ 1214 "PSE_T≔pose_trans(pose_inv(FRM_Reference), CAM_OBJ_Pose)"
            global PSE_T= pose_trans ( pose_inv (FRM_Reference), CAM_OBJ_Pose)
            $ 1215 "CAM_Result.append(get_pattern_counter(PSE_T, 'X', pattern=[10, 5], patternsize=[0.181, 0.081]))"
            CAM_Result.append(get_pattern_counter(PSE_T, "X", pattern=[10, 5], patternsize=[0.181, 0.081]))
            $ 1216 "PRC_CntDetect≔PRC_CntDetect+1"
            global PRC_CntDetect=PRC_CntDetect+1
          end
          $ 1217 "CAM_Done≔ True "
          global CAM_Done=  True
        else:
          $ 1218 "ElseIf CAM_Captures≥CAM_PRM_Retries"
          if (CAM_Captures >= CAM_PRM_Retries):
            $ 1219 "CAM_Done≔ True "
            global CAM_Done=  True
          else:
            $ 1220 "Else" "noBreak"
            $ 1221 "CAM_Captures≔CAM_Captures+1"
            global CAM_Captures=CAM_Captures+1
          end
        end
      end
    end
    $ 1222 "'=========='"
    # '=========='
    $ 1223 "PostSettings"
    $ 1224 "FRM_Reference≔p[0,0,0,0,0,0]"
    global FRM_Reference=p[0,0,0,0,0,0]
    $ 1225 "Set"
    set_tcp(p[0.0,0.0,0.161,3.1415,0.0,0.0])
    $ 1226 "CAM_Pose≔p[0,0,0,0,0,0]"
    global CAM_Pose=p[0,0,0,0,0,0]
    $ 1227 "Action≔0"
    global Action=0
    $ 1228 "Action_Info≔''"
    global Action_Info=""
  end
  def Sub_AMR_MiR_V3():
    $ 1229 "Sub_AMR_MiR_V3" "noBreak"
    $ 1230 "PreSettings"
    $ 1231 "AMR_TargetList≔[1,2,3,4,5,21,22,23,24,31,32,33,34,35,36,37,38,41]"
    global AMR_TargetList=[1,2,3,4,5,21,22,23,24,31,32,33,34,35,36,37,38,41]
    $ 1232 "AMR_Done≔ False "
    global AMR_Done=  False
    $ 1233 "AMR_PosActual≔T2O_Current_Pos"
    global AMR_PosActual=modbus_get_signal_status("T2O_Current_Pos")
    $ 1234 "AMR_Attemps≔T2O_Nav_Attemps"
    global AMR_Attemps=modbus_get_signal_status("T2O_Nav_Attemps")
    $ 1235 "AMR_Battery≔MiR_Battery_Lvl"
    global AMR_Battery=modbus_get_signal_status("MiR_Battery_Lvl")
    $ 1236 "AMR_Charging≔(T2O_Charging≟1)"
    global AMR_Charging=(modbus_get_signal_status("T2O_Charging") == 1)
    $ 1237 "AMR_Position≔struct(position_identifier=T2O_Current_Pos, x1=MiR_Position_X1, x2=MiR_Position_X2, y1=MiR_Position_Y1, y2=MiR_Position_Y2, theta1=MiR_Theta_1, theta2=MiR_Theta_2) "
    global AMR_Position=struct(position_identifier=modbus_get_signal_status("T2O_Current_Pos"), x1=modbus_get_signal_status("MiR_Position_X1"), x2=modbus_get_signal_status("MiR_Position_X2"), y1=modbus_get_signal_status("MiR_Position_Y1"), y2=modbus_get_signal_status("MiR_Position_Y2"), theta1=modbus_get_signal_status("MiR_Theta_1"), theta2=modbus_get_signal_status("MiR_Theta_2"))
    $ 1238 "If MiR_Mode≠7"
    if (modbus_get_signal_status("MiR_Mode") != 7):
      $ 1239 "Error"
      $ 1240 "set_error(ERROR_AMR_WRONG_MODE)"
      set_error(ERROR_AMR_WRONG_MODE)
      $ 1241 "AMR_Done≔ True "
      global AMR_Done=  True
    end
    $ 1242 "'=========='"
    # '=========='
    $ 1243 "Switch STATE"
    switch_1 = STATE
    $ 1244 "Case 1"
    if (1 == switch_1):
      $ 1245 "stopping"
      $ 1246 "If T2O_Done≟1 and O2T_Acknowledge≟0"
      if (modbus_get_signal_status("T2O_Done") == 1  and  modbus_get_signal_status("O2T_Acknowledge") == 0):
        $ 1247 "Set O2T_Acknowledge=1"
        modbus_set_output_register("O2T_Acknowledge", 1)
      end
      $ 1248 "Set MiR_CMD_Stop=On"
      modbus_set_output_signal("MiR_CMD_Stop", True)
      $ 1249 "AMR_Position.position_identifier = 0"
      AMR_Position.position_identifier = 0
      $ 1250 "AMR_Done≔ True "
      global AMR_Done=  True
    elif (2 == switch_1):
      $ 1251 "Case 2"
      $ 1252 "stopped"
      $ 1253 "If MiR_State≠3 and MiR_State≠5"
      if (modbus_get_signal_status("MiR_State") != 3  and  modbus_get_signal_status("MiR_State") != 5):
        $ 1254 "Set MiR_CMD_Stop=Off"
        modbus_set_output_signal("MiR_CMD_Stop", False)
      end
    elif (3 == switch_1):
      $ 1255 "Case 3"
      $ 1256 "resetting"
      $ 1257 "Set O2T_Mis_Main=Off"
      modbus_set_output_signal("O2T_Mis_Main", False)
      $ 1258 "Set O2T_Mis_Charge=Off"
      modbus_set_output_signal("O2T_Mis_Charge", False)
      $ 1259 "If MiR_Mis_Queue>0"
      if (modbus_get_signal_status("MiR_Mis_Queue")>0):
        $ 1260 "Set MiR_CMD_Clear_Q=On"
        modbus_set_output_signal("MiR_CMD_Clear_Q", True)
        $ 1261 "Wait MiR_Mis_Queue≟0"
        while (not(modbus_get_signal_status("MiR_Mis_Queue") == 0)):
          sync()
        end
        $ 1262 "Set MiR_CMD_Clear_Q=Off"
        modbus_set_output_signal("MiR_CMD_Clear_Q", False)
      end
      $ 1263 "If MiR_Error_ID≠0"
      if (modbus_get_signal_status("MiR_Error_ID") != 0):
        $ 1264 "Set MiR_CMD_Clear_E=On"
        modbus_set_output_signal("MiR_CMD_Clear_E", True)
        $ 1265 "Wait MiR_Error_ID≟0"
        while (not(modbus_get_signal_status("MiR_Error_ID") == 0)):
          sync()
        end
        $ 1266 "Set MiR_CMD_Clear_E=Off"
        modbus_set_output_signal("MiR_CMD_Clear_E", False)
      end
      $ 1267 "Set O2T_Action=0"
      modbus_set_output_register("O2T_Action", 0)
      $ 1268 "Set O2T_Acknowledge=0"
      modbus_set_output_register("O2T_Acknowledge", 0)
      $ 1269 "Set O2T_Target_Pos=0"
      modbus_set_output_register("O2T_Target_Pos", 0)
      $ 1270 "Set O2T_Footprint=0"
      modbus_set_output_register("O2T_Footprint", 0)
      $ 1271 "Set O2T_ProtectOff=0"
      modbus_set_output_register("O2T_ProtectOff", 0)
      $ 1272 "Set O2T_Dock=0"
      modbus_set_output_register("O2T_Dock", 0)
      $ 1273 "AMR_Attemps≔0"
      global AMR_Attemps=0
      $ 1274 "AMR_PosTarget≔0"
      global AMR_PosTarget=0
      $ 1275 "AMR_Step≔0"
      global AMR_Step=0
      $ 1276 "AMR_AtTarget≔ False "
      global AMR_AtTarget=  False
      $ 1277 "If MiR_State≟4 or MiR_State≟3 or MiR_State≟10"
      if (modbus_get_signal_status("MiR_State") == 4  or  modbus_get_signal_status("MiR_State") == 3  or  modbus_get_signal_status("MiR_State") == 10):
        $ 1278 "AMR_Done≔ True "
        global AMR_Done=  True
      end
    elif (5 == switch_1):
      $ 1279 "Case 5"
      $ 1280 "starting"
      $ 1281 "If MiR_State≟4"
      if (modbus_get_signal_status("MiR_State") == 4):
        $ 1282 "Set MiR_CMD_Start=On"
        modbus_set_output_signal("MiR_CMD_Start", True)
        $ 1283 "Wait MiR_State≠4"
        while (not(modbus_get_signal_status("MiR_State") != 4)):
          sync()
        end
        $ 1284 "Set MiR_CMD_Start=Off"
        modbus_set_output_signal("MiR_CMD_Start", False)
        $ 1285 "AMR_Done≔ True "
        global AMR_Done=  True
      else:
        $ 1286 "ElseIf MiR_State≟10"
        if (modbus_get_signal_status("MiR_State") == 10):
          $ 1287 "'MiR in protective stop. Wait'"
          # 'MiR in protective stop. Wait'
          $ 1288 "AMR_Done≔ True "
          global AMR_Done=  True
        else:
          $ 1289 "ElseIf MiR_State≟3"
          if (modbus_get_signal_status("MiR_State") == 3):
            $ 1290 "AMR_Done≔ True "
            global AMR_Done=  True
          end
        end
      end
    elif (6 == switch_1):
      $ 1291 "Case 6"
      $ 1292 "execute"
      $ 1293 "AMR_AtTarget≔(AMR_PosActual≟AMR_PosTarget)"
      global AMR_AtTarget=(AMR_PosActual == AMR_PosTarget)
      $ 1294 "Switch AMR_Step"
      switch_2 = AMR_Step
      $ 1295 "Case 0"
      if (0 == switch_2):
        $ 1296 "If  not AMR_AtTarget"
        if (  not  AMR_AtTarget):
          $ 1297 "AMR_Step≔1"
          global AMR_Step=1
        else:
          $ 1298 "Else" "noBreak"
          $ 1299 "AMR_Done≔ True "
          global AMR_Done=  True
        end
      elif (1 == switch_2):
        $ 1300 "Case 1"
        $ 1301 "general Settings"
        $ 1302 "Set O2T_Acknowledge=0"
        modbus_set_output_register("O2T_Acknowledge", 0)
        $ 1303 "check for error"
        $ 1304 "If OBJ_Picked and MiR_State≟10"
        if (OBJ_Picked  and  modbus_get_signal_status("MiR_State") == 10):
          $ 1305 "Error"
          $ 1306 "set_error(ERROR_ROBOT_ARM_NOT_IN_HOME_POSE)"
          set_error(ERROR_ROBOT_ARM_NOT_IN_HOME_POSE)
          $ 1307 "Action≔0"
          global Action=0
        else:
          $ 1308 "ElseIf  not found_in_list(AMR_PosTarget, AMR_TargetList)"
          if (  not  found_in_list(AMR_PosTarget, AMR_TargetList)):
            $ 1309 "Error"
            $ 1310 "set_error(ERROR_UNKNOWN_POSE)"
            set_error(ERROR_UNKNOWN_POSE)
            $ 1311 "Action≔0"
            global Action=0
          end
        end
        $ 1312 "If MiR_State≟3"
        if (modbus_get_signal_status("MiR_State") == 3):
          $ 1313 "Set MiR_CMD_Start=Off"
          modbus_set_output_signal("MiR_CMD_Start", False)
          $ 1314 "Switch Action"
          switch_3 = Action
          $ 1315 "Case 51"
          if (51 == switch_3):
            $ 1316 "Charge"
            $ 1317 "'trigger the charging mission'"
            # 'trigger the charging mission'
            $ 1318 "'target pos is predefined'"
            # 'target pos is predefined'
            $ 1319 "Set O2T_Footprint=0"
            modbus_set_output_register("O2T_Footprint", 0)
            $ 1320 "Set O2T_Action=1"
            modbus_set_output_register("O2T_Action", 1)
            $ 1321 "If MiR_Mis_Queue≟0"
            if (modbus_get_signal_status("MiR_Mis_Queue") == 0):
              $ 1322 "Set O2T_Mis_Charge=On"
              modbus_set_output_signal("O2T_Mis_Charge", True)
              $ 1323 "Wait MiR_Mis_Queue≥1"
              while (not(modbus_get_signal_status("MiR_Mis_Queue") >= 1)):
                sync()
              end
              $ 1324 "Set O2T_Mis_Charge=Off"
              modbus_set_output_signal("O2T_Mis_Charge", False)
            end
          elif (52 == switch_3):
            $ 1325 "Case 52"
            $ 1326 "Navigate"
            $ 1327 "'trigger the standard missoin'"
            # 'trigger the standard missoin'
            $ 1328 "Set O2T_Footprint=AMR_FootprintID"
            modbus_set_output_register("O2T_Footprint", AMR_FootprintID)
            $ 1329 "Set O2T_Target_Pos=AMR_PosTarget"
            modbus_set_output_register("O2T_Target_Pos", AMR_PosTarget)
            $ 1330 "Set O2T_Action=2"
            modbus_set_output_register("O2T_Action", 2)
            $ 1331 "If MiR_Mis_Queue≟0"
            if (modbus_get_signal_status("MiR_Mis_Queue") == 0):
              $ 1332 "Set O2T_Mis_Main=On"
              modbus_set_output_signal("O2T_Mis_Main", True)
              $ 1333 "Wait MiR_Mis_Queue≥1"
              while (not(modbus_get_signal_status("MiR_Mis_Queue") >= 1)):
                sync()
              end
              $ 1334 "Set O2T_Mis_Main=Off"
              modbus_set_output_signal("O2T_Mis_Main", False)
            end
          end
        else:
          $ 1335 "ElseIf MiR_State≟4"
          if (modbus_get_signal_status("MiR_State") == 4):
            $ 1336 "Set MiR_CMD_Start=On"
            modbus_set_output_signal("MiR_CMD_Start", True)
          else:
            $ 1337 "ElseIf MiR_State≟5"
            if (modbus_get_signal_status("MiR_State") == 5):
              $ 1338 "AMR_Step≔2"
              global AMR_Step=2
            else:
              $ 1339 "ElseIf MiR_State≟10"
              if (modbus_get_signal_status("MiR_State") == 10):
                $ 1340 "'AMR still in safeguard stop'"
                # 'AMR still in safeguard stop'
              end
            end
          end
        end
      elif (2 == switch_2):
        $ 1341 "Case 2"
        $ 1342 "acknowledge handshake"
        $ 1343 "If T2O_Done≟1 and O2T_Acknowledge≟0"
        if (modbus_get_signal_status("T2O_Done") == 1  and  modbus_get_signal_status("O2T_Acknowledge") == 0):
          $ 1344 "Set O2T_Acknowledge=1"
          modbus_set_output_register("O2T_Acknowledge", 1)
        else:
          $ 1345 "ElseIf T2O_Done≟0 and O2T_Acknowledge≟1"
          if (modbus_get_signal_status("T2O_Done") == 0  and  modbus_get_signal_status("O2T_Acknowledge") == 1):
            $ 1346 "Set O2T_Acknowledge=0"
            modbus_set_output_register("O2T_Acknowledge", 0)
            $ 1347 "AMR_AtTarget≔(AMR_PosActual≟AMR_PosTarget)"
            global AMR_AtTarget=(AMR_PosActual == AMR_PosTarget)
            $ 1348 "AMR_Done≔ True "
            global AMR_Done=  True
          end
        end
      end
      $ 1349 "translate errors"
      $ 1350 "If AMR_Done"
      if (AMR_Done):
        $ 1351 "Switch T2O_Error_ID"
        switch_2 = modbus_get_signal_status("T2O_Error_ID")
        $ 1352 "Case 2003"
        if (2003 == switch_2):
          $ 1353 "error"
          $ 1354 "set_error(ERROR_NOT_DOCKED)"
          set_error(ERROR_NOT_DOCKED)
        elif (2007 == switch_2):
          $ 1355 "Case 2007"
          $ 1356 "error"
          $ 1357 "set_error(ERROR_NOT_REACHABLE_TARGET)"
          set_error(ERROR_NOT_REACHABLE_TARGET)
        elif (2008 == switch_2):
          $ 1358 "Case 2008"
          $ 1359 "error"
          $ 1360 "set_error(ERROR_CHARGING_NOT_STARTED)"
          set_error(ERROR_CHARGING_NOT_STARTED)
        end
      end
    elif (7 == switch_1):
      $ 1361 "Case 7"
      $ 1362 "completing"
      $ 1363 "If MiR_Mis_Queue>0"
      if (modbus_get_signal_status("MiR_Mis_Queue")>0):
        $ 1364 "Set MiR_CMD_Abort=On"
        modbus_set_output_signal("MiR_CMD_Abort", True)
        $ 1365 "Wait MiR_Mis_Queue≟0"
        while (not(modbus_get_signal_status("MiR_Mis_Queue") == 0)):
          sync()
        end
        $ 1366 "Set MiR_CMD_Abort=Off"
        modbus_set_output_signal("MiR_CMD_Abort", False)
      end
      $ 1367 "If MiR_State≟3 or MiR_State≟10"
      if (modbus_get_signal_status("MiR_State") == 3  or  modbus_get_signal_status("MiR_State") == 10):
        $ 1368 "AMR_Done≔ True "
        global AMR_Done=  True
      end
    elif (9 == switch_1):
      $ 1369 "Case 9"
      $ 1370 "holding"
      $ 1371 "Set MiR_CMD_Abort=On"
      modbus_set_output_signal("MiR_CMD_Abort", True)
      $ 1372 "If MiR_State≟3 or MiR_State≟10"
      if (modbus_get_signal_status("MiR_State") == 3  or  modbus_get_signal_status("MiR_State") == 10):
        $ 1373 "Set MiR_CMD_Abort=Off"
        modbus_set_output_signal("MiR_CMD_Abort", False)
        $ 1374 "AMR_Done≔ True "
        global AMR_Done=  True
      end
    elif (11 == switch_1):
      $ 1375 "Case 11"
      $ 1376 "unholding"
      $ 1377 "Set MiR_CMD_Start=On"
      modbus_set_output_signal("MiR_CMD_Start", True)
      $ 1378 "If MiR_State≠4"
      if (modbus_get_signal_status("MiR_State") != 4):
        $ 1379 "Set MiR_CMD_Start=Off"
        modbus_set_output_signal("MiR_CMD_Start", False)
        $ 1380 "AMR_Step≔0"
        global AMR_Step=0
        $ 1381 "AMR_Done≔ True "
        global AMR_Done=  True
      end
    elif (12 == switch_1):
      $ 1382 "Case 12"
      $ 1383 "suspending"
      $ 1384 "'none'"
      # 'none'
    elif (14 == switch_1):
      $ 1385 "Case 14"
      $ 1386 "unsuspending"
      $ 1387 "'none'"
      # 'none'
    elif (15 == switch_1):
      $ 1388 "Case 15"
      $ 1389 "aborting"
      $ 1390 "Set MiR_CMD_Abort=On"
      modbus_set_output_signal("MiR_CMD_Abort", True)
      $ 1391 "Wait MiR_State≟3"
      while (not(modbus_get_signal_status("MiR_State") == 3)):
        sync()
      end
      $ 1392 "Set MiR_CMD_Abort=Off"
      modbus_set_output_signal("MiR_CMD_Abort", False)
    elif (17 == switch_1):
      $ 1393 "Case 17"
      $ 1394 "clearing"
      $ 1395 "If MiR_Error_ID≠0"
      if (modbus_get_signal_status("MiR_Error_ID") != 0):
        $ 1396 "Set MiR_CMD_Clear_E=On"
        modbus_set_output_signal("MiR_CMD_Clear_E", True)
        $ 1397 "Wait MiR_Error_ID≟0"
        while (not(modbus_get_signal_status("MiR_Error_ID") == 0)):
          sync()
        end
        $ 1398 "Set MiR_CMD_Clear_E=Off"
        modbus_set_output_signal("MiR_CMD_Clear_E", False)
      end
      $ 1399 "If MiR_Error_ID≟0"
      if (modbus_get_signal_status("MiR_Error_ID") == 0):
        $ 1400 "AMR_Done≔ True "
        global AMR_Done=  True
      end
    end
    $ 1401 "'=========='"
    # '=========='
    $ 1402 "PostSettings"
    $ 1403 "AMR_Position≔struct(position_identifier=T2O_Current_Pos, x1=MiR_Position_X1, x2=MiR_Position_X2, y1=MiR_Position_Y1, y2=MiR_Position_Y2, theta1=MiR_Theta_1, theta2=MiR_Theta_2) "
    global AMR_Position=struct(position_identifier=modbus_get_signal_status("T2O_Current_Pos"), x1=modbus_get_signal_status("MiR_Position_X1"), x2=modbus_get_signal_status("MiR_Position_X2"), y1=modbus_get_signal_status("MiR_Position_Y1"), y2=modbus_get_signal_status("MiR_Position_Y2"), theta1=modbus_get_signal_status("MiR_Theta_1"), theta2=modbus_get_signal_status("MiR_Theta_2"))
  end
  def Sub_Action_V4():
    $ 1404 "Sub_Action_V4" "noBreak"
    $ 1405 "PreSettings"
    $ 1406 "init poses"
    $ 1407 "PSE_A≔p[0,0,0,0,0,0]"
    global PSE_A=p[0,0,0,0,0,0]
    $ 1408 "PSE_A_H≔p[0,0,0,0,0,0]"
    global PSE_A_H=p[0,0,0,0,0,0]
    $ 1409 "PSE_T≔p[0,0,0,0,0,0]"
    global PSE_T=p[0,0,0,0,0,0]
    $ 1410 "PSE_T_H≔p[0,0,0,0,0,0]"
    global PSE_T_H=p[0,0,0,0,0,0]
    $ 1411 "PSE_G≔p[0,0,0,0,0,0]"
    global PSE_G=p[0,0,0,0,0,0]
    $ 1412 "PSE_G_H≔p[0,0,0,0,0,0]"
    global PSE_G_H=p[0,0,0,0,0,0]
    $ 1413 "PSE_R≔p[0,0,0,0,0,0]"
    global PSE_R=p[0,0,0,0,0,0]
    $ 1414 "PSE_R_H≔p[0,0,0,0,0,0]"
    global PSE_R_H=p[0,0,0,0,0,0]
    $ 1415 "JNT_Q≔[0,0,0,0,0,0]"
    global JNT_Q=[0,0,0,0,0,0]
    $ 1416 "JNT_S≔[0,0,0,0,0,0]"
    global JNT_S=[0,0,0,0,0,0]
    $ 1417 "Gripping parameters"
    $ 1418 "OBJ = find_object_by_type(OBJs, OBJ_Type)"
    OBJ = find_object_by_type(OBJs, OBJ_Type)
    $ 1419 "GRP_Open_Pos≔OBJ.dimension.diameter * 1000 + 6"
    global GRP_Open_Pos=OBJ.dimension.diameter * 1000 + 6
    $ 1420 "GRP_Offset≔OBJ.gripper_offset"
    global GRP_Offset=OBJ.gripper_offset
    $ 1421 "rq_set_force_norm(50)"
     rq_set_force_norm (50)
    $ 1422 "rq_set_speed_norm(50)"
     rq_set_speed_norm (50)
    $ 1423 "Switch ITM_ID"
    switch_1 = ITM_ID
    $ 1424 "Case 1"
    if (1 == switch_1):
      $ 1425 "uML"
      $ 1426 "JIG2 = find_object_by_type(JIGs, JIG)"
      JIG2 = find_object_by_type(JIGs, JIG)
      $ 1427 "JIG_Offset≔JIG2.jig_offset"
      global JIG_Offset=JIG2.jig_offset
      $ 1428 "Switch JIG"
      switch_2 = JIG
      $ 1429 "Case 1"
      if (1 == switch_2):
        $ 1430 "3FG"
        $ 1431 "define poses"
        $ 1432 "FRM_Reference≔ULM_3FG"
        global FRM_Reference=ULM_3FG
        $ 1433 "JNT_Q≔JNT_HOME"
        global JNT_Q=JNT_HOME
        $ 1434 "PSE_T≔pose_trans(GRP_Offset, JIG_Offset)"
        global PSE_T= pose_trans (GRP_Offset, JIG_Offset)
        $ 1435 "PSE_A≔pose_trans(PSE_T, p[0,0,0.100,0,0,0])"
        global PSE_A= pose_trans (PSE_T, p[0,0,0.100,0,0,0])
        $ 1436 "PSE_R≔pose_add(PSE_T, p[0,0,0.100,0,0,0])"
        global PSE_R= pose_add (PSE_T, p[0,0,0.100,0,0,0])
      elif (2 == switch_2):
        $ 1437 "Case 2"
        $ 1438 "Input"
        $ 1439 "'CHANGE THE REFERENCE TO THE FRAME TO MOVE IN'"
        # 'CHANGE THE REFERENCE TO THE FRAME TO MOVE IN'
        $ 1440 "define poses"
        $ 1441 "FRM_Reference≔ULM_Input"
        global FRM_Reference=ULM_Input
        $ 1442 "PSE_T≔pose_trans(pose_trans(get_pattern_pos_rectangle(OBJ_Nbr, 'X', [10,5], patternsize=[0.181,0.081]), GRP_Offset), JIG_Offset)"
        global PSE_T= pose_trans ( pose_trans (get_pattern_pos_rectangle(OBJ_Nbr, "X", [10,5], patternsize=[0.181,0.081]), GRP_Offset), JIG_Offset)
        $ 1443 "If Action≟1"
        if (Action == 1):
          $ 1444 "PSE_R≔pose_add(PSE_T, p[0,0,0.200,0,0,0])"
          global PSE_R= pose_add (PSE_T, p[0,0,0.200,0,0,0])
          $ 1445 "PSE_A≔pose_add(PSE_T, p[0,0,0.100,0,0,0])"
          global PSE_A= pose_add (PSE_T, p[0,0,0.100,0,0,0])
        else:
          $ 1446 "ElseIf Action≟2"
          if (Action == 2):
            $ 1447 "PSE_R≔pose_add(PSE_T, p[0,0,0.100,0,0,0])"
            global PSE_R= pose_add (PSE_T, p[0,0,0.100,0,0,0])
            $ 1448 "PSE_A≔pose_add(PSE_T, p[0,0,0.200,0,0,0])"
            global PSE_A= pose_add (PSE_T, p[0,0,0.200,0,0,0])
          end
        end
      elif (3 == switch_2):
        $ 1449 "Case 3"
        $ 1450 "Output"
        $ 1451 "'CHANGE THE REFERENCE TO THE FRAME TO MOVE IN'"
        # 'CHANGE THE REFERENCE TO THE FRAME TO MOVE IN'
        $ 1452 "define poses"
        $ 1453 "FRM_Reference≔ULM_Output"
        global FRM_Reference=ULM_Output
        $ 1454 "PSE_T≔pose_trans(pose_trans(get_pattern_pos_rectangle(OBJ_Nbr, 'X', [10,5], patternsize=[0.181,0.081]), GRP_Offset), JIG_Offset)"
        global PSE_T= pose_trans ( pose_trans (get_pattern_pos_rectangle(OBJ_Nbr, "X", [10,5], patternsize=[0.181,0.081]), GRP_Offset), JIG_Offset)
        $ 1456 "If Action≟1"
        if (Action == 1):
          $ 1457 "PSE_R≔pose_add(PSE_T, p[0,0,0.200,0,0,0])"
          global PSE_R= pose_add (PSE_T, p[0,0,0.200,0,0,0])
          $ 1458 "PSE_A≔pose_add(PSE_T, p[0,0,0.100,0,0,0])"
          global PSE_A= pose_add (PSE_T, p[0,0,0.100,0,0,0])
        else:
          $ 1459 "ElseIf Action≟2"
          if (Action == 2):
            $ 1460 "PSE_R≔pose_add(PSE_T, p[0,0,0.100,0,0,0])"
            global PSE_R= pose_add (PSE_T, p[0,0,0.100,0,0,0])
            $ 1461 "PSE_A≔pose_add(PSE_T, p[0,0,0.200,0,0,0])"
            global PSE_A= pose_add (PSE_T, p[0,0,0.200,0,0,0])
          end
        end
      elif (4 == switch_2):
        $ 1462 "Case 4"
        $ 1463 "jig centrifuge racks"
        $ 1464 "define poses"
        $ 1465 "FRM_Reference≔ULM_Cent_Racks"
        global FRM_Reference=ULM_Cent_Racks
        $ 1466 "PSE_T≔get_pattern_pos_rectangle(JIG_Slot, 'X', [4,1], patternsize=[0.291,0])"
        global PSE_T=get_pattern_pos_rectangle(JIG_Slot, "X", [4,1], patternsize=[0.291,0])
        $ 1467 "If OBJ_Nbr≠0"
        if (OBJ_Nbr != 0):
          $ 1468 "PSE_T≔pose_trans(pose_trans(PSE_T, get_pattern_pos_rectangle(OBJ_Nbr, 'X', [3,3], patternsize=[0.060,0.060])),p[-0.030, -0.030,0,0,0,3.927])"
          global PSE_T= pose_trans ( pose_trans (PSE_T, get_pattern_pos_rectangle(OBJ_Nbr, "X", [3,3], patternsize=[0.060,0.060])),p[-0.030, -0.030,0,0,0,3.927])
        end
        $ 1469 "PSE_T≔pose_trans(PSE_T, GRP_Offset)"
        global PSE_T= pose_trans (PSE_T, GRP_Offset)
        $ 1470 "If Action≟1"
        if (Action == 1):
          $ 1471 "PSE_R≔pose_add(PSE_T, p[0,0,0.200,0,0,0])"
          global PSE_R= pose_add (PSE_T, p[0,0,0.200,0,0,0])
          $ 1472 "PSE_A≔pose_add(PSE_T, p[0,0,0.100,0,0,0])"
          global PSE_A= pose_add (PSE_T, p[0,0,0.100,0,0,0])
        else:
          $ 1473 "ElseIf Action≟2"
          if (Action == 2):
            $ 1474 "PSE_R≔pose_add(PSE_T, p[0,0,0.100,0,0,0])"
            global PSE_R= pose_add (PSE_T, p[0,0,0.100,0,0,0])
            $ 1475 "PSE_A≔pose_add(PSE_T, p[0,0,0.200,0,0,0])"
            global PSE_A= pose_add (PSE_T, p[0,0,0.200,0,0,0])
          end
        end
      elif (6 == switch_2):
        $ 1476 "Case 6"
        $ 1477 "Caps bin"
        $ 1478 "define poses"
        $ 1479 "'Drop cap'"
        # 'Drop cap'
        $ 1480 "FRM_Reference=ULM_Cap_Bin"
        FRM_Reference=ULM_Cap_Bin
        $ 1481 "PSE_T≔pose_RPY2RotVec(p[0,0,0,0,0,0])"
        global PSE_T=pose_RPY2RotVec(p[0,0,0,0,0,0])
        $ 1482 "PSE_T_H≔pose_add(PSE_T, p[0,0,-0.011,0,0,0])"
        global PSE_T_H= pose_add (PSE_T, p[0,0,-0.011,0,0,0])
        $ 1483 "PSE_A≔pose_trans(PSE_T, p[0,0,0.1,0,0,0])"
        global PSE_A= pose_trans (PSE_T, p[0,0,0.1,0,0,0])
        $ 1484 "PSE_R_H≔pose_add(PSE_T, p[0,0,0.100,0,0,0])"
        global PSE_R_H= pose_add (PSE_T, p[0,0,0.100,0,0,0])
        $ 1485 "PSE_R≔pose_add(PSE_T, p[0,0,0.100,0,0,0])"
        global PSE_R= pose_add (PSE_T, p[0,0,0.100,0,0,0])
      elif (7 == switch_2):
        $ 1486 "Case 7"
        $ 1487 "Sarstedt"
        $ 1488 "'CHANGE THE REFERENCE TO THE FRAME TO MOVE IN'"
        # 'CHANGE THE REFERENCE TO THE FRAME TO MOVE IN'
        $ 1494 "If TASK.ID≟10"
        if (TASK.ID == 10):
          $ 1495 "Frame & Position Params"
          $ 1497 "FRM_Reference = CAM_LM_SSRack"
          FRM_Reference = CAM_LM_SSRack
          $ 1502 "PSE_T≔uLM_SS_PickPlc"
          global PSE_T=uLM_SS_PickPlc
          $ 1503 "PSE_A≔pose_trans(PSE_T, p[0,0,0.1,0,0,0])"
          global PSE_A= pose_trans (PSE_T, p[0,0,0.1,0,0,0])
          $ 1504 "PSE_R≔pose_add(PSE_T, p[0,0,0.1,0,0,0])"
          global PSE_R= pose_add (PSE_T, p[0,0,0.1,0,0,0])
        else:
          $ 1505 "ElseIf TASK.ID≟11"
          if (TASK.ID == 11):
            $ 1506 "FRM_Reference = ULM_SS_Jig"
            FRM_Reference = ULM_SS_Jig
            $ 1507 "PSE_T≔pose_RPY2RotVec(p[0,0,0,0,0,0])"
            global PSE_T=pose_RPY2RotVec(p[0,0,0,0,0,0])
            $ 1508 "PSE_T≔pose_trans(PSE_T, GRP_Offset)"
            global PSE_T=pose_trans(PSE_T, GRP_Offset)
            $ 1509 "PSE_A≔pose_trans(PSE_T, p[0,0,0.1,0,0,0])"
            global PSE_A= pose_trans (PSE_T, p[0,0,0.1,0,0,0])
            $ 1510 "PSE_R≔pose_add(PSE_T, p[0,0,0.2,0,0,0])"
            global PSE_R= pose_add (PSE_T, p[0,0,0.2,0,0,0])
          end
        end
      elif (8 == switch_2):
        $ 1511 "Case 8"
        $ 1512 "NoK"
        $ 1513 "define poses"
        $ 1514 "'NoK'"
        # 'NoK'
        $ 1515 "FRM_Reference=ULM_NoK"
        FRM_Reference=ULM_NoK
        $ 1516 "PSE_T≔pose_RPY2RotVec(p[0,0,0,0,0,0])"
        global PSE_T=pose_RPY2RotVec(p[0,0,0,0,0,0])
        $ 1517 "PSE_A≔pose_trans(PSE_T, p[0,0,0.1,0,0,0])"
        global PSE_A= pose_trans (PSE_T, p[0,0,0.1,0,0,0])
        $ 1518 "PSE_R≔pose_add(PSE_T, p[0,0,0.100,0,0,0])"
        global PSE_R= pose_add (PSE_T, p[0,0,0.100,0,0,0])
      elif (9 == switch_2):
        $ 1519 "Case 9"
      elif (10 == switch_2):
        $ 1527 "Case 10"
      elif (11 == switch_2):
        $ 1535 "Case 11"
      elif (12 == switch_2):
        $ 1543 "Case 12"
      end
    elif (2 == switch_1):
      $ 1551 "Case 2"
      $ 1552 "Centrifuge"
      $ 1553 "'CHANGE THE REFERENCE TO THE FRAME TO MOVE IN'"
      # 'CHANGE THE REFERENCE TO THE FRAME TO MOVE IN'
      $ 1554 "define poses"
      $ 1555 "FRM_Reference≔FRM_Centrifuge"
      global FRM_Reference=FRM_Centrifuge
      $ 1556 "PSE_T≔GRP_Offset"
      global PSE_T=GRP_Offset
      $ 1557 "If Action≟8"
      if (Action == 8):
        $ 1558 "PSE_R≔pose_add(PSE_T, p[0,0,0.250,0,0,0])"
        global PSE_R= pose_add (PSE_T, p[0,0,0.250,0,0,0])
        $ 1559 "PSE_A≔pose_add(PSE_T, p[0,0,0.150,0,0,0])"
        global PSE_A= pose_add (PSE_T, p[0,0,0.150,0,0,0])
      else:
        $ 1560 "ElseIf Action≟7"
        if (Action == 7):
          $ 1561 "PSE_R≔pose_add(PSE_T, p[0,0,0.150,0,0,0])"
          global PSE_R= pose_add (PSE_T, p[0,0,0.150,0,0,0])
          $ 1562 "PSE_A≔pose_add(PSE_T, p[0,0,0.250,0,0,0])"
          global PSE_A= pose_add (PSE_T, p[0,0,0.250,0,0,0])
        end
      end
    elif (3 == switch_1):
      $ 1563 "Case 3"
      $ 1564 "Output"
      $ 1565 "'CHANGE THE REFERENCE TO THE FRAME TO MOVE IN'"
      # 'CHANGE THE REFERENCE TO THE FRAME TO MOVE IN'
      $ 1566 "define poses"
      $ 1567 "FRM_Reference≔Base_const"
      global FRM_Reference=p[0.0,0.0,0.0,0.0,0.0,0.0]
      $ 1568 "PSE_T≔p[0,0,0,0,0,0]"
      global PSE_T=p[0,0,0,0,0,0]
      $ 1569 "PSE_A≔pose_add(PSE_T, p[0,0,0.150,0,0,0])"
      global PSE_A= pose_add (PSE_T, p[0,0,0.150,0,0,0])
      $ 1570 "PSE_R≔pose_add(PSE_T, p[0,0,0.100,0,0,0])"
      global PSE_R= pose_add (PSE_T, p[0,0,0.100,0,0,0])
    elif (5 == switch_1):
      $ 1571 "Case 5"
      $ 1572 "Sarstedt Pickup Table"
      $ 1573 "'CHANGE THE REFERENCE TO THE FRAME TO MOVE IN'"
      # 'CHANGE THE REFERENCE TO THE FRAME TO MOVE IN'
      $ 1574 "Switch JIG"
      switch_2 = JIG
      $ 1575 "Case 7"
      if (7 == switch_2):
        $ 1588 "Sarstedt"
        $ 1589 "'CHANGE THE REFERENCE TO THE FRAME TO MOVE IN'"
        # 'CHANGE THE REFERENCE TO THE FRAME TO MOVE IN'
        $ 1595 "If TASK.ID≟10"
        if (TASK.ID == 10):
          $ 1596 "Frame & Position Params"
          $ 1597 "FRM_Reference = CAM_LM_SSRack"
          FRM_Reference = CAM_LM_SSRack
          $ 1598 "PSE_T≔uLM_SS_PickPlc"
          global PSE_T=uLM_SS_PickPlc
          $ 1599 "PSE_A≔pose_trans(PSE_T, p[0,0,0.1,0,0,0])"
          global PSE_A= pose_trans (PSE_T, p[0,0,0.1,0,0,0])
          $ 1600 "PSE_R≔pose_add(PSE_T, p[0,0,0.1,0,0,0])"
          global PSE_R= pose_add (PSE_T, p[0,0,0.1,0,0,0])
        end
      end
    elif (13 == switch_1):
      $ 1607 "Case 13"
      $ 1608 "Sarstedt Pickup Table"
      $ 1609 "'CHANGE THE REFERENCE TO THE FRAME TO MOVE IN'"
      # 'CHANGE THE REFERENCE TO THE FRAME TO MOVE IN'
      $ 1610 "Switch JIG"
      switch_2 = JIG
      $ 1611 "Case 7"
      if (7 == switch_2):
        $ 1624 "Bottle"
        $ 1625 "'CHANGE THE REFERENCE TO THE FRAME TO MOVE IN'"
        # 'CHANGE THE REFERENCE TO THE FRAME TO MOVE IN'
        $ 1631 "If TASK.ID≟43"
        if (TASK.ID == 43):
          $ 1632 "Frame & Position Params"
          $ 1634 "PSE_T≔uLM_SS_PickPlc"
          global PSE_T=uLM_SS_PickPlc
          $ 1635 "PSE_A≔pose_trans(PSE_T, p[0,0,0.1,0,0,0])"
          global PSE_A= pose_trans (PSE_T, p[0,0,0.1,0,0,0])
          $ 1636 "PSE_R≔pose_add(PSE_T, p[0,0,0.1,0,0,0])"
          global PSE_R= pose_add (PSE_T, p[0,0,0.1,0,0,0])
        end
      end
    end
    $ 1643 "Additional check"
    $ 1644 "If  not is_reachable(FRM_Reference,[PSE_A,PSE_A_H,PSE_T,PSE_T_H,PSE_R,PSE_R_H])"
    if (  not  is_reachable(FRM_Reference,[PSE_A,PSE_A_H,PSE_T,PSE_T_H,PSE_R,PSE_R_H])):
      $ 1645 "Error"
      $ 1646 "set_error(ERROR_POSE_NOT_REACHABLE)"
      set_error(ERROR_POSE_NOT_REACHABLE)
      $ 1647 "Action≔0"
      global Action=0
    end
    $ 1648 "'=========='"
    # '=========='
    $ 1649 "Switch Action"
    switch_1 = Action
    $ 1650 "Case 1"
    if (1 == switch_1):
      $ 1651 "Pick"
      $ 1652 "Action_Info≔'pick object'"
      global Action_Info="pick object"
      $ 1653 "do_transition(pose_trans(FRM_Reference, PSE_T), keep_rxry=OBJ_Picked)"
      do_transition( pose_trans (FRM_Reference, PSE_T), keep_rxry=OBJ_Picked)
      $ 1654 "EOAT"
      $ 1655 "If  not OBJ_Picked"
      if (  not  OBJ_Picked):
        $ 1656 "rq_move_and_wait_mm(GRP_Open_Pos)"
         rq_move_and_wait_mm (GRP_Open_Pos)
      end
      $ 1657 "If PSE_A_H≠PSE_Z"
      if (PSE_A_H != PSE_Z):
        $ 1658 "If JNT_Q≠JNT_Z"
        if (JNT_Q != JNT_Z):
          $ 1659 "movej(get_inverse_kin(pose_trans(FRM_Reference, PSE_A_H), qnear=JNT_Q), r=0.050)"
          movej(get_inverse_kin( pose_trans (FRM_Reference, PSE_A_H), qnear=JNT_Q), r=0.050)
        else:
          $ 1660 "Else" "noBreak"
          $ 1661 "movej(pose_trans(FRM_Reference, PSE_A_H), r=0.050)"
          movej( pose_trans (FRM_Reference, PSE_A_H), r=0.050)
        end
      end
      $ 1662 "If PSE_A≠PSE_Z"
      if (PSE_A != PSE_Z):
        $ 1663 "If JNT_Q≠JNT_Z"
        if (JNT_Q != JNT_Z):
          $ 1664 "movej(get_inverse_kin(pose_trans(FRM_Reference, PSE_A), qnear=JNT_Q), r=0.020)"
          movej(get_inverse_kin( pose_trans (FRM_Reference, PSE_A), qnear=JNT_Q), r=0.020)
        else:
          $ 1665 "Else" "noBreak"
          $ 1666 "movej(pose_trans(FRM_Reference, PSE_A), r=0.020)"
          movej( pose_trans (FRM_Reference, PSE_A), r=0.020)
        end
      end
      $ 1667 "MoveL"
      $ 1668 "If PSE_T_H≠PSE_Z"
      if (PSE_T_H != PSE_Z):
        $ 1669 "PSE_T_H" "breakAfter"
        movel(pose_trans(FRM_Reference, PSE_T_H), a=0.5, v=0.4, r=0.01)
      end
      $ 1670 "PSE_T" "breakAfter"
      movel(pose_trans(FRM_Reference, PSE_T), a=0.08, v=0.12)
      $ 1671 "EOAT"
      $ 1672 "rq_set_force_norm(50)"
       rq_set_force_norm (50)
      $ 1673 "rq_close_and_wait()"
       rq_close_and_wait ()
      $ 1674 "OBJ_Picked≔rq_is_object_detected()"
      global OBJ_Picked= rq_is_object_detected ()
      $ 1675 "If  not OBJ_Picked"
      if (  not  OBJ_Picked):
        $ 1676 "set_error(ERROR_NO_OBJECT_TO_PICK)"
        set_error(ERROR_NO_OBJECT_TO_PICK)
      end
      $ 1677 "EXTT"
      $ 1678 "Switch JIG"
      switch_2 = JIG
      $ 1679 "Case 1"
      if (1 == switch_2):
        $ 1680 "3FG"
        $ 1681 "If OBJ_Picked"
        if (OBJ_Picked):
          $ 1682 "Set GRP_3F_Open=On"
          set_standard_digital_out(5, True)
        end
      end
      $ 1683 "If PSE_R_H≠PSE_Z"
      if (PSE_R_H != PSE_Z):
        $ 1684 "PSE_R" "breakAfter"
        movel(pose_trans(FRM_Reference, PSE_R), a=0.5, v=0.4, r=0.01)
        $ 1685 "PSE_R_H" "breakAfter"
        movel(pose_trans(FRM_Reference, PSE_R_H), a=0.5, v=0.4)
      else:
        $ 1686 "Else" "noBreak"
        $ 1687 "PSE_R" "breakAfter"
        movel(pose_trans(FRM_Reference, PSE_R), a=0.5, v=0.4)
      end
    elif (2 == switch_1):
      $ 1688 "Case 2"
      $ 1689 "Place"
      $ 1690 "Action_Info≔'place object'"
      global Action_Info="place object"
      $ 1691 "do_transition(pose_trans(FRM_Reference, PSE_T), keep_rxry=OBJ_Picked)"
      do_transition( pose_trans (FRM_Reference, PSE_T), keep_rxry=OBJ_Picked)
      $ 1692 "EXTT"
      $ 1693 "Switch JIG"
      switch_2 = JIG
      $ 1694 "Case 1"
      if (1 == switch_2):
        $ 1695 "3FG"
        $ 1696 "If OBJ_Picked"
        if (OBJ_Picked):
          $ 1697 "Set GRP_3F_Open=On"
          set_standard_digital_out(5, True)
        end
      end
      $ 1698 "If PSE_A_H≠PSE_Z"
      if (PSE_A_H != PSE_Z):
        $ 1699 "If JNT_Q≠JNT_Z"
        if (JNT_Q != JNT_Z):
          $ 1700 "movej(get_inverse_kin(pose_trans(FRM_Reference, PSE_A_H), qnear=JNT_Q), r=0.050)"
          movej(get_inverse_kin( pose_trans (FRM_Reference, PSE_A_H), qnear=JNT_Q), r=0.050)
        else:
          $ 1701 "Else" "noBreak"
          $ 1702 "movej(pose_trans(FRM_Reference, PSE_A_H), r=0.050)"
          movej( pose_trans (FRM_Reference, PSE_A_H), r=0.050)
        end
      end
      $ 1703 "If PSE_A≠PSE_Z"
      if (PSE_A != PSE_Z):
        $ 1704 "If JNT_Q≠JNT_Z"
        if (JNT_Q != JNT_Z):
          $ 1705 "movej(get_inverse_kin(pose_trans(FRM_Reference, PSE_A), qnear=JNT_Q), r=0.020)"
          movej(get_inverse_kin( pose_trans (FRM_Reference, PSE_A), qnear=JNT_Q), r=0.020)
        else:
          $ 1706 "Else" "noBreak"
          $ 1707 "movej(pose_trans(FRM_Reference, PSE_A), r=0.020)"
          movej( pose_trans (FRM_Reference, PSE_A), r=0.020)
        end
      end
      $ 1708 "MoveL"
      $ 1709 "If PSE_T_H≠PSE_Z"
      if (PSE_T_H != PSE_Z):
        $ 1710 "PSE_T_H" "breakAfter"
        movel(pose_trans(FRM_Reference, PSE_T_H), a=0.5, v=0.4, r=0.01)
      end
      $ 1711 "PSE_T" "breakAfter"
      global move_thread_flag_1711=0
      thread move_thread_1711():
        enter_critical
        move_thread_flag_1711 = 1
        movel(pose_trans(FRM_Reference, PSE_T), a=0.05, v=0.09)
        move_thread_flag_1711 = 2
        exit_critical
      end
      move_thread_flag_1711 = 0
      move_thread_han_1711 = run move_thread_1711()
      while (True):
        local targetTcpDirection=get_target_tcp_speed()
        local stepsToRetract=tool_contact(direction=targetTcpDirection)
        if (stepsToRetract > 0):
          kill move_thread_han_1711
          stopl(0.5)
          $ 1712 "Until (tool_contact_detection)"
          break
        end
        sleep(1.0E-10)
        if (move_thread_flag_1711 > 1):
          join move_thread_han_1711
          break
        end
        sync()
      end
      $ 1713 "Force"
      sleep(0.02)
      zero_ftsensor()
      force_mode(FRM_Reference, [1, 1, 1, 0, 0, 0], [0.0, 0.0, 0.0, 0.0, 0.0, 0.0], 2, [0.1, 0.1, 0.01, 0.3490658503988659, 0.3490658503988659, 0.3490658503988659])
      $ 1714 "PSE_T" "noBreak"
      movel(pose_trans(FRM_Reference, PSE_T), a=0.04, v=0.07)
      end_force_mode()
      stopl(5.0)
      $ 1715 "EXTT"
      $ 1716 "Switch JIG"
      switch_2 = JIG
      $ 1717 "Case 1"
      if (1 == switch_2):
        $ 1718 "3FG"
        $ 1719 "If OBJ_Picked"
        if (OBJ_Picked):
          $ 1720 "Set GRP_3F_Open=Off"
          set_standard_digital_out(5, False)
          $ 1721 "Wait: 0.2"
          sleep(0.2)
        end
      end
      $ 1722 "EOAT"
      $ 1723 "rq_move_and_wait_mm(GRP_Open_Pos)"
       rq_move_and_wait_mm (GRP_Open_Pos)
      $ 1724 "OBJ_Picked≔rq_is_object_detected()"
      global OBJ_Picked= rq_is_object_detected ()
      $ 1725 "If PSE_R_H≠PSE_Z"
      if (PSE_R_H != PSE_Z):
        $ 1726 "PSE_R" "breakAfter"
        movel(pose_trans(FRM_Reference, PSE_R), a=0.5, v=0.4, r=0.01)
        $ 1727 "PSE_R_H" "breakAfter"
        movel(pose_trans(FRM_Reference, PSE_R_H), a=0.5, v=0.4)
      else:
        $ 1728 "Else" "noBreak"
        $ 1729 "PSE_R" "breakAfter"
        movel(pose_trans(FRM_Reference, PSE_R), a=0.5, v=0.4)
      end
    elif (3 == switch_1):
      $ 1730 "Case 3"
      $ 1731 "Push"
      $ 1732 "Action_Info≔'push'"
      global Action_Info="push"
    elif (4 == switch_1):
      $ 1733 "Case 4"
      $ 1734 "Pull"
      $ 1735 "Action_Info≔'pull'"
      global Action_Info="pull"
    elif (6 == switch_1):
      $ 1738 "Case 6"
      $ 1739 "Drop the cap"
      $ 1740 "If JNT_A≠[0,0,0,0,0,0]"
      if (JNT_A != [0,0,0,0,0,0]):
        $ 1741 "MoveJ"
        $ 1742 "JNT_A" "breakAfter"
        movej(JNT_A, a=1.3962634015954636, v=1.7453292519943295, r=0.02)
      else:
        $ 1743 "Else" "noBreak"
        $ 1744 "MoveJ"
        $ 1745 "PSE_A" "breakAfter"
        movej(pose_trans(FRM_Reference, PSE_A), a=1.3962634015954636, v=1.7453292519943295, r=0.02)
      end
      $ 1746 "MoveL"
      $ 1747 "PSE_T" "breakAfter"
      movel(pose_trans(FRM_Reference, PSE_T), a=0.05, v=0.09)
      $ 1748 "'ADD OPEN GRIPPER'"
      # 'ADD OPEN GRIPPER'
      # begin: URCap Program Node
      #   Source: Robotiq_Grippers, 3.17.0.105337, Robotiq Inc.
      #   Type: Gripper
      $ 1749 "Gripper Move10mm (1)"
      if not(gripper_connected[0]):
        popup("Gripper 1 must be connected to run this program.", "No connection", False, True, True)
      end
      if not(rq_is_gripper_activated("1")):
        popup("Gripper 1 is not activated. Go to Installation tab > Gripper to activate it and run the program again.", "Not activated", False, True, True)
      end
      rq_set_pos_spd_for(201, 0, 28, "1")
      rq_wait_pos_spe_for_request(201, 0, 28, "1")
      rq_go_to("1")
      rq_wait("1")
      # end: URCap Program Node
      $ 1750 "PSE_T_H" "breakAfter"
      movel(pose_trans(FRM_Reference, PSE_T_H), a=0.05, v=0.09)
      # begin: URCap Program Node
      #   Source: Robotiq_Grippers, 3.17.0.105337, Robotiq Inc.
      #   Type: Gripper
      $ 1751 "Gripper Move40mm (1)"
      if not(gripper_connected[0]):
        popup("Gripper 1 must be connected to run this program.", "No connection", False, True, True)
      end
      if not(rq_is_gripper_activated("1")):
        popup("Gripper 1 is not activated. Go to Installation tab > Gripper to activate it and run the program again.", "Not activated", False, True, True)
      end
      rq_set_pos_spd_for(63, 0, 28, "1")
      rq_wait_pos_spe_for_request(63, 0, 28, "1")
      rq_go_to("1")
      rq_wait("1")
      # end: URCap Program Node
      $ 1752 "PSE_R" "breakAfter"
      movel(pose_trans(FRM_Reference, PSE_R), a=0.5, v=0.4)
    elif (7 == switch_1):
      $ 1753 "Case 7"
      $ 1754 "Load"
      $ 1755 "Action_Info≔'load object'"
      global Action_Info="load object"
      $ 1756 "do_transition(pose_trans(FRM_Reference, PSE_T), keep_rxry=OBJ_Picked)"
      do_transition( pose_trans (FRM_Reference, PSE_T), keep_rxry=OBJ_Picked)
      $ 1757 "If PSE_A_H≠PSE_Z"
      if (PSE_A_H != PSE_Z):
        $ 1758 "If JNT_Q≠JNT_Z"
        if (JNT_Q != JNT_Z):
          $ 1759 "movej(get_inverse_kin(pose_trans(FRM_Reference, PSE_A_H), qnear=JNT_Q), r=0.050)"
          movej(get_inverse_kin( pose_trans (FRM_Reference, PSE_A_H), qnear=JNT_Q), r=0.050)
        else:
          $ 1760 "Else" "noBreak"
          $ 1761 "movej(pose_trans(FRM_Reference, PSE_A_H), r=0.050)"
          movej( pose_trans (FRM_Reference, PSE_A_H), r=0.050)
        end
      end
      $ 1762 "If PSE_A≠PSE_Z"
      if (PSE_A != PSE_Z):
        $ 1763 "If JNT_Q≠JNT_Z"
        if (JNT_Q != JNT_Z):
          $ 1764 "movej(get_inverse_kin(pose_trans(FRM_Reference, PSE_A), qnear=JNT_Q), r=0.020)"
          movej(get_inverse_kin( pose_trans (FRM_Reference, PSE_A), qnear=JNT_Q), r=0.020)
        else:
          $ 1765 "Else" "noBreak"
          $ 1766 "movej(pose_trans(FRM_Reference, PSE_A), r=0.020)"
          movej( pose_trans (FRM_Reference, PSE_A), r=0.020)
        end
      end
      $ 1767 "MoveL"
      $ 1768 "If PSE_T_H≠PSE_Z"
      if (PSE_T_H != PSE_Z):
        $ 1769 "PSE_T_H" "breakAfter"
        movel(pose_trans(FRM_Reference, PSE_T_H), a=0.5, v=0.4, r=0.01)
      end
      $ 1770 "PSE_T" "breakAfter"
      global move_thread_flag_1770=0
      thread move_thread_1770():
        enter_critical
        move_thread_flag_1770 = 1
        movel(pose_trans(FRM_Reference, PSE_T), a=0.05, v=0.09)
        move_thread_flag_1770 = 2
        exit_critical
      end
      move_thread_flag_1770 = 0
      move_thread_han_1770 = run move_thread_1770()
      while (True):
        local targetTcpDirection=get_target_tcp_speed()
        local stepsToRetract=tool_contact(direction=targetTcpDirection)
        if (stepsToRetract > 0):
          kill move_thread_han_1770
          stopl(0.5)
          $ 1771 "Until (tool_contact_detection)"
          break
        end
        sleep(1.0E-10)
        if (move_thread_flag_1770 > 1):
          join move_thread_han_1770
          break
        end
        sync()
      end
      $ 1772 "Force"
      sleep(0.02)
      zero_ftsensor()
      force_mode(FRM_Reference, [0, 1, 1, 0, 0, 1], [0.0, 0.0, 0.0, 0.0, 0.0, 0.0], 2, [0.1, 0.05, 0.02, 0.3490658503988659, 0.3490658503988659, 3.141592653589793])
      $ 1773 "PSE_T" "noBreak"
      movel(pose_trans(FRM_Reference, PSE_T), a=0.04, v=0.07)
      end_force_mode()
      stopl(5.0)
      $ 1774 "EOAT"
      $ 1775 "rq_move_and_wait_mm(GRP_Open_Pos)"
       rq_move_and_wait_mm (GRP_Open_Pos)
      $ 1776 "OBJ_Picked≔rq_is_object_detected()"
      global OBJ_Picked= rq_is_object_detected ()
      $ 1777 "If PSE_R_H≠PSE_Z"
      if (PSE_R_H != PSE_Z):
        $ 1778 "PSE_R" "breakAfter"
        movel(pose_trans(FRM_Reference, PSE_R), a=0.5, v=0.4, r=0.01)
        $ 1779 "PSE_R_H" "breakAfter"
        movel(pose_trans(FRM_Reference, PSE_R_H), a=0.5, v=0.4)
      else:
        $ 1780 "Else" "noBreak"
        $ 1781 "PSE_R" "breakAfter"
        movel(pose_trans(FRM_Reference, PSE_R), a=0.5, v=0.4)
      end
    elif (8 == switch_1):
      $ 1782 "Case 8"
      $ 1783 "Unload"
      $ 1784 "Action_Info≔'pick object'"
      global Action_Info="pick object"
      $ 1785 "do_transition(pose_trans(FRM_Reference, PSE_T), keep_rxry=OBJ_Picked)"
      do_transition( pose_trans (FRM_Reference, PSE_T), keep_rxry=OBJ_Picked)
      $ 1786 "EOAT"
      $ 1787 "If  not OBJ_Picked"
      if (  not  OBJ_Picked):
        $ 1788 "rq_move_and_wait_mm(GRP_Open_Pos)"
         rq_move_and_wait_mm (GRP_Open_Pos)
      end
      $ 1789 "If PSE_A_H≠PSE_Z"
      if (PSE_A_H != PSE_Z):
        $ 1790 "If JNT_Q≠JNT_Z"
        if (JNT_Q != JNT_Z):
          $ 1791 "movej(get_inverse_kin(pose_trans(FRM_Reference, PSE_A_H), qnear=JNT_Q), r=0.050)"
          movej(get_inverse_kin( pose_trans (FRM_Reference, PSE_A_H), qnear=JNT_Q), r=0.050)
        else:
          $ 1792 "Else" "noBreak"
          $ 1793 "movej(pose_trans(FRM_Reference, PSE_A_H), r=0.050)"
          movej( pose_trans (FRM_Reference, PSE_A_H), r=0.050)
        end
      end
      $ 1794 "If PSE_A≠PSE_Z"
      if (PSE_A != PSE_Z):
        $ 1795 "If JNT_Q≠JNT_Z"
        if (JNT_Q != JNT_Z):
          $ 1796 "movej(get_inverse_kin(pose_trans(FRM_Reference, PSE_A), qnear=JNT_Q), r=0.020)"
          movej(get_inverse_kin( pose_trans (FRM_Reference, PSE_A), qnear=JNT_Q), r=0.020)
        else:
          $ 1797 "Else" "noBreak"
          $ 1798 "movej(pose_trans(FRM_Reference, PSE_A), r=0.020)"
          movej( pose_trans (FRM_Reference, PSE_A), r=0.020)
        end
      end
      $ 1799 "MoveL"
      $ 1800 "If PSE_T_H≠PSE_Z"
      if (PSE_T_H != PSE_Z):
        $ 1801 "PSE_T_H" "breakAfter"
        movel(pose_trans(FRM_Reference, PSE_T_H), a=0.5, v=0.4, r=0.01)
      end
      $ 1802 "PSE_T" "breakAfter"
      movel(pose_trans(FRM_Reference, PSE_T), a=0.08, v=0.12)
      $ 1803 "Force"
      sleep(0.02)
      zero_ftsensor()
      force_mode(FRM_Reference, [1, 1, 0, 0, 0, 0], [0.0, 0.0, 0.0, 0.0, 0.0, 0.0], 2, [0.05, 0.05, 0.1, 0.3490658503988659, 0.3490658503988659, 0.3490658503988659])
      $ 1804 "EOAT" "noBreak"
      $ 1805 "rq_set_force_norm(50)" "noBreak"
       rq_set_force_norm (50)
      $ 1806 "rq_close_and_wait()" "noBreak"
       rq_close_and_wait ()
      $ 1807 "OBJ_Picked≔rq_is_object_detected()" "noBreak"
      global OBJ_Picked= rq_is_object_detected ()
      $ 1808 "If  not OBJ_Picked" "noBreak"
      if (  not  OBJ_Picked):
        $ 1809 "set_error(ERROR_NO_OBJECT_TO_PICK)" "noBreak"
        set_error(ERROR_NO_OBJECT_TO_PICK)
      end
      $ 1810 "If PSE_R_H≠PSE_Z" "noBreak"
      if (PSE_R_H != PSE_Z):
        $ 1811 "PSE_R" "noBreak"
        movel(pose_trans(FRM_Reference, PSE_R), a=0.5, v=0.4, r=0.01)
        $ 1812 "PSE_R_H" "noBreak"
        movel(pose_trans(FRM_Reference, PSE_R_H), a=0.5, v=0.4)
      else:
        $ 1813 "Else" "noBreak"
        $ 1814 "PSE_R" "noBreak"
        movel(pose_trans(FRM_Reference, PSE_R), a=0.5, v=0.4)
      end
      end_force_mode()
      stopl(5.0)
    elif (11 == switch_1):
      $ 1815 "Case 11"
    elif (12 == switch_1):
      $ 1852 "Case 12"
      $ 1853 "Decap"
      $ 1854 "Action_Info≔'decapping'"
      global Action_Info="decapping"
      $ 1855 "Set GRP_3F_Enable=On"
      set_standard_digital_out(4, True)
      $ 1856 "Set GRP_3F_Decap=On"
      set_standard_digital_out(3, True)
      $ 1857 "Force"
      sleep(0.02)
      zero_ftsensor()
      force_mode(tool_pose(), [0, 0, 1, 0, 0, 0], [0.0, 0.0, 5.0, 0.0, 0.0, 0.0], 2, [0.1, 0.1, 0.15, 0.3490658503988659, 0.3490658503988659, 0.3490658503988659])
      $ 1858 "check_decapping(offset=0.015, timeout=5, abort=CMD_Hold)" "noBreak"
      check_decapping(offset=0.015, timeout=5, abort=CMD_Hold)
      end_force_mode()
      stopl(5.0)
      $ 1859 "Set GRP_3F_Decap=Off"
      set_standard_digital_out(3, False)
      $ 1860 "Set GRP_3F_Enable=Off"
      set_standard_digital_out(4, False)
      $ 1861 "MoveL"
      $ 1862 "PSE_R" "breakAfter"
      movel(pose_trans(FRM_Reference, PSE_R), a=0.8, v=0.15)
    elif (13 == switch_1):
      $ 1863 "Case 13"
      $ 1864 "TMR_Barcode: Reset"
      TMR_Barcode = 0
      $ 1865 "Read"
      $ 1866 "TMR_Barcode: Start"
      TMR_Barcode_is_counting = True
      $ 1867 "If TMR_Barcode<PRM_TO_Read_BC"
      global thread_flag_1867=0
      thread Thread_if_1867():
        $ 1868 "KeyenceTrigger"
        $ 1869 "Set OClearResult=HI:Pulse 0.2"
        thread SinglePulse18():
          write_output_boolean_register(2, True)
          sleep(0.2)
          write_output_boolean_register(2, False)
        end
        singlePulse18 = run SinglePulse18()
        $ 1870 "Wait: 0.5"
        sleep(0.5)
        $ 1871 "Set OTriggerBarcode=Off"
        write_output_boolean_register(1, False)
        $ 1872 "Wait: 0.5"
        sleep(0.5)
        $ 1873 "Set OTriggerBarcode=On"
        write_output_boolean_register(1, True)
        $ 1874 "Wait: 0.5"
        sleep(0.5)
        $ 1875 "Preorient"
        $ 1876 "TMR_Barcode: Reset"
        TMR_Barcode = 0
        $ 1877 "If ICmdExctd"
        if (read_input_boolean_register(12)):
          $ 1878 "Set GRP_3F_Decap=On"
          set_standard_digital_out(3, True)
          $ 1879 "Set GRP_3F_Enable=On"
          set_standard_digital_out(4, True)
          $ 1880 "Loop ICmdExctd"
          while (read_input_boolean_register(12)):
            $ 1881 "KeyenceTrigger"
            $ 1882 "Set OClearResult=HI:Pulse 0.1"
            thread SinglePulse19():
              write_output_boolean_register(2, True)
              sleep(0.1)
              write_output_boolean_register(2, False)
            end
            singlePulse19 = run SinglePulse19()
            $ 1883 "Wait: 0.3"
            sleep(0.3)
            $ 1884 "Set OTriggerBarcode=Off"
            write_output_boolean_register(1, False)
            $ 1885 "Wait: 0.3"
            sleep(0.3)
            $ 1886 "Set OTriggerBarcode=On"
            write_output_boolean_register(1, True)
            $ 1887 "Wait: 0.1"
            sleep(0.1)
          end
        end
        $ 1888 "If  not ICmdExctd"
        if (  not  read_input_boolean_register(12)):
          $ 1889 "Set GRP_3F_Decap=On"
          set_standard_digital_out(3, True)
          $ 1890 "Set GRP_3F_Enable=On"
          set_standard_digital_out(4, True)
          $ 1891 "Wait ICmdExctd=HI"
          while (read_input_boolean_register(12) == False):
            sync()
          end
        end
        $ 1892 "Set GRP_3F_Decap=Off"
        set_standard_digital_out(3, False)
        $ 1893 "Set GRP_3F_Enable=Off"
        set_standard_digital_out(4, False)
        $ 1894 "OBJ_Brc_OK≔ True "
        global OBJ_Brc_OK=  True
        thread_flag_1867 = 1
      end
      if (TMR_Barcode<PRM_TO_Read_BC):
        global thread_handler_1867=run Thread_if_1867()
        while (thread_flag_1867 == 0):
          if not(TMR_Barcode<PRM_TO_Read_BC):
            kill thread_handler_1867
            thread_flag_1867 = 2
          else:
            sync()
          end
        end
      else:
        thread_flag_1867 = 2
      end
      if (thread_flag_1867 == 2):
        $ 1895 "Else" "noBreak"
        $ 1896 "exeption"
        $ 1897 "error"
        $ 1899 "OBJ_Brc_OK≔ False "
        global OBJ_Brc_OK=  False
      end
      $ 1900 "Set GRP_3F_Decap=Off"
      set_standard_digital_out(3, False)
      $ 1901 "Set GRP_3F_Enable=Off"
      set_standard_digital_out(4, False)
      $ 1902 "Set OTriggerBarcode=Off"
      write_output_boolean_register(1, False)
    elif (15 == switch_1):
      $ 1903 "Case 15"
      $ 1904 "Detect"
      $ 1905 "Action_Info≔'detect'"
      global Action_Info="detect"
    elif (30 == switch_1):
      $ 1906 "Case 30"
      $ 1907 "Shake"
      $ 1908 "Action_Info≔'shake'"
      global Action_Info="shake"
      $ 1909 "do_transition(pose_trans(FRM_Reference, PSE_T), keep_rxry=OBJ_Picked)"
      do_transition( pose_trans (FRM_Reference, PSE_T), keep_rxry=OBJ_Picked)
      $ 1910 "If PSE_A_H≠PSE_Z"
      if (PSE_A_H != PSE_Z):
        $ 1911 "If JNT_Q≠JNT_Z"
        if (JNT_Q != JNT_Z):
          $ 1912 "movej(get_inverse_kin(pose_trans(FRM_Reference, PSE_A_H), qnear=JNT_Q), r=0.050)"
          movej(get_inverse_kin( pose_trans (FRM_Reference, PSE_A_H), qnear=JNT_Q), r=0.050)
        else:
          $ 1913 "Else" "noBreak"
          $ 1914 "movej(pose_trans(FRM_Reference, PSE_A_H), r=0.050)"
          movej( pose_trans (FRM_Reference, PSE_A_H), r=0.050)
        end
      end
      $ 1915 "If PSE_A≠PSE_Z"
      if (PSE_A != PSE_Z):
        $ 1916 "If JNT_Q≠JNT_Z"
        if (JNT_Q != JNT_Z):
          $ 1917 "movej(get_inverse_kin(pose_trans(FRM_Reference, PSE_A), qnear=JNT_Q), r=0.020)"
          movej(get_inverse_kin( pose_trans (FRM_Reference, PSE_A), qnear=JNT_Q), r=0.020)
        else:
          $ 1918 "Else" "noBreak"
          $ 1919 "movej(pose_trans(FRM_Reference, PSE_A), r=0.020)"
          movej( pose_trans (FRM_Reference, PSE_A), r=0.020)
        end
      end
      $ 1920 "MoveL"
      $ 1921 "If PSE_T_H≠PSE_Z"
      if (PSE_T_H != PSE_Z):
        $ 1922 "PSE_T_H" "breakAfter"
        movel(pose_trans(FRM_Reference, PSE_T_H), a=0.5, v=0.4, r=0.01)
      end
      $ 1923 "PSE_T" "breakAfter"
